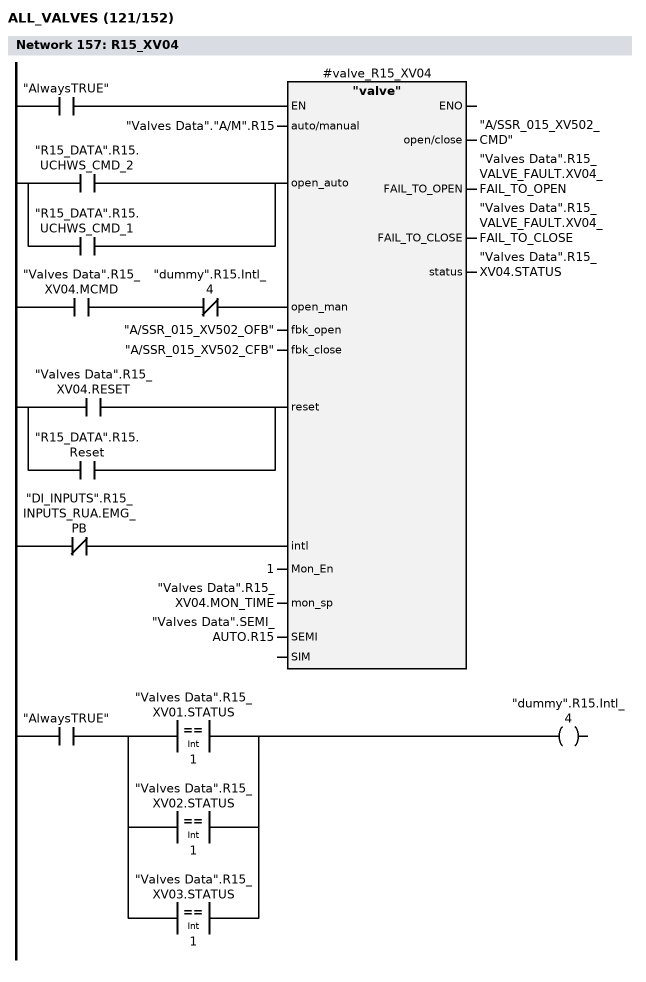
   RUNG wire#powerrail
      Contact( "AlwaysTRUE" )
      #valve_R15_XV04(open_auto := wire#w1, open_man := wire#w2, reset := wire#w3, intl := wire#w4, "auto/manual" := "Valves Data"."A/M".R15, fbk_open := "A/SSR_015_XV502_OFB", fbk_close := "A/SSR_015_XV502_CFB", Mon_En := 1, mon_sp := "Valves Data".R15_XV04.MON_TIME, SEMI := "Valves Data".SEMI_AUTO.R15, SIM :=, "open/close" => "A/SSR_015_XV502_CMD", FAIL_TO_OPEN => "Valves Data".R15_VALVE_FAULT.XV04_FAIL_TO_OPEN, FAIL_TO_CLOSE => "Valves Data".R15_VALVE_FAULT.XV04_FAIL_TO_CLOSE, status => "Valves Data".R15_XV04.STATUS)
   END_RUNG
   RUNG wire#powerrail
      Contact( "R15_DATA".R15.UCHWS_CMD_2 )
   END_RUNG wire#w1
   RUNG wire#powerrail
      Contact( "R15_DATA".R15.UCHWS_CMD_1 )
   END_RUNG wire#w1
   RUNG wire#powerrail
      Contact( "Valves Data".R15_XV04.MCMD )
      I_Contact( "dummy".R15.Intl_4 )
   END_RUNG wire#w2
   RUNG wire#powerrail
      Contact( "Valves Data".R15_XV04.RESET )
   END_RUNG wire#w3
   RUNG wire#powerrail
      Contact( "R15_DATA".R15.Reset )
   END_RUNG wire#w3
   RUNG wire#powerrail
      I_Contact( "DI_INPUTS".R15_INPUTS_RUA.EMG_PB )
   END_RUNG wire#w4
   RUNG wire#powerrail
      Contact( "AlwaysTRUE" )
      wire#w5
      { S7_Templates := "SrcType := Int" } EQ_Contact(in1 := "Valves Data".R15_XV01.STATUS, in2 := 1)
      wire#w6
      Coil( "dummy".R15.Intl_4 )
   END_RUNG
   RUNG wire#w5
      { S7_Templates := "SrcType := Int" } EQ_Contact(in1 := "Valves Data".R15_XV02.STATUS, in2 := 1)
   END_RUNG wire#w6
   RUNG wire#w5
      { S7_Templates := "SrcType := Int" } EQ_Contact(in1 := "Valves Data".R15_XV03.STATUS, in2 := 1)
   END_RUNG wire#w6
   // the same network as SCL:
   IF "AlwaysTRUE" THEN
       #valve_R15_XV04("auto/manual" := "Valves Data"."A/M".R15,   // "valve"
                       open_auto := "R15_DATA".R15.UCHWS_CMD_2 OR "R15_DATA".R15.UCHWS_CMD_1,
                       open_man := "Valves Data".R15_XV04.MCMD AND NOT "dummy".R15.Intl_4,
                       fbk_open := "A/SSR_015_XV502_OFB",
                       fbk_close := "A/SSR_015_XV502_CFB",
                       reset := "Valves Data".R15_XV04.RESET OR "R15_DATA".R15.Reset,
                       intl := NOT "DI_INPUTS".R15_INPUTS_RUA.EMG_PB,
                       Mon_En := 1,
                       mon_sp := "Valves Data".R15_XV04.MON_TIME,
                       SEMI := "Valves Data".SEMI_AUTO.R15,
                       "open/close" => "A/SSR_015_XV502_CMD",
                       FAIL_TO_OPEN => "Valves Data".R15_VALVE_FAULT.XV04_FAIL_TO_OPEN,
                       FAIL_TO_CLOSE => "Valves Data".R15_VALVE_FAULT.XV04_FAIL_TO_CLOSE,
                       status => "Valves Data".R15_XV04.STATUS);
   END_IF;
   "dummy".R15.Intl_4 := "AlwaysTRUE" AND (("Valves Data".R15_XV01.STATUS = 1) OR ("Valves Data".R15_XV02.STATUS = 1) OR ("Valves Data".R15_XV03.STATUS = 1));
END_REGION

REGION Network 158: R15_XV05
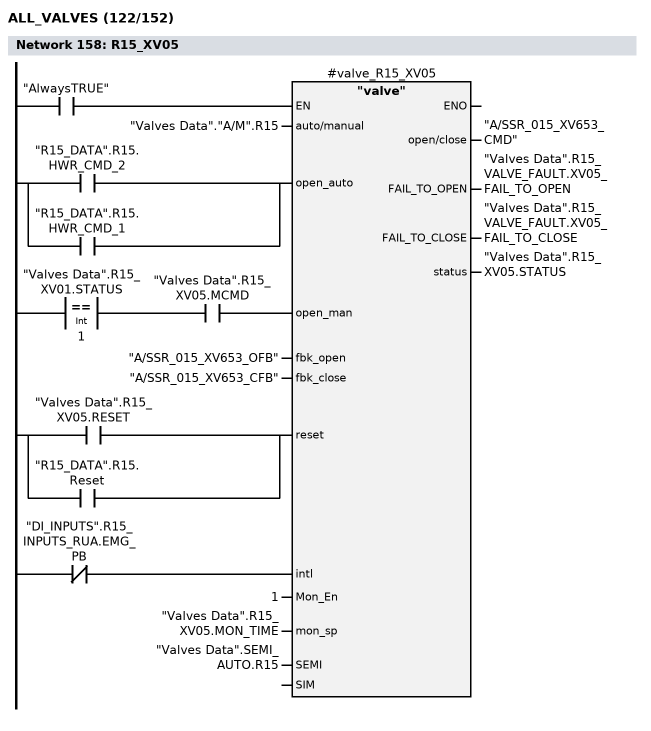
   RUNG wire#powerrail
      Contact( "AlwaysTRUE" )
      #valve_R15_XV05(open_auto := wire#w1, open_man := wire#w2, reset := wire#w3, intl := wire#w4, "auto/manual" := "Valves Data"."A/M".R15, fbk_open := "A/SSR_015_XV653_OFB", fbk_close := "A/SSR_015_XV653_CFB", Mon_En := 1, mon_sp := "Valves Data".R15_XV05.MON_TIME, SEMI := "Valves Data".SEMI_AUTO.R15, SIM :=, "open/close" => "A/SSR_015_XV653_CMD", FAIL_TO_OPEN => "Valves Data".R15_VALVE_FAULT.XV05_FAIL_TO_OPEN, FAIL_TO_CLOSE => "Valves Data".R15_VALVE_FAULT.XV05_FAIL_TO_CLOSE, status => "Valves Data".R15_XV05.STATUS)
   END_RUNG
   RUNG wire#powerrail
      Contact( "R15_DATA".R15.HWR_CMD_2 )
   END_RUNG wire#w1
   RUNG wire#powerrail
      Contact( "R15_DATA".R15.HWR_CMD_1 )
   END_RUNG wire#w1
   RUNG wire#powerrail
      { S7_Templates := "SrcType := Int" } EQ_Contact(in1 := "Valves Data".R15_XV01.STATUS, in2 := 1)
      Contact( "Valves Data".R15_XV05.MCMD )
   END_RUNG wire#w2
   RUNG wire#powerrail
      Contact( "Valves Data".R15_XV05.RESET )
   END_RUNG wire#w3
   RUNG wire#powerrail
      Contact( "R15_DATA".R15.Reset )
   END_RUNG wire#w3
   RUNG wire#powerrail
      I_Contact( "DI_INPUTS".R15_INPUTS_RUA.EMG_PB )
   END_RUNG wire#w4
   // the same network as SCL:
   IF "AlwaysTRUE" THEN
       #valve_R15_XV05("auto/manual" := "Valves Data"."A/M".R15,   // "valve"
                       open_auto := "R15_DATA".R15.HWR_CMD_2 OR "R15_DATA".R15.HWR_CMD_1,
                       open_man := ("Valves Data".R15_XV01.STATUS = 1) AND "Valves Data".R15_XV05.MCMD,
                       fbk_open := "A/SSR_015_XV653_OFB",
                       fbk_close := "A/SSR_015_XV653_CFB",
                       reset := "Valves Data".R15_XV05.RESET OR "R15_DATA".R15.Reset,
                       intl := NOT "DI_INPUTS".R15_INPUTS_RUA.EMG_PB,
                       Mon_En := 1,
                       mon_sp := "Valves Data".R15_XV05.MON_TIME,
                       SEMI := "Valves Data".SEMI_AUTO.R15,
                       "open/close" => "A/SSR_015_XV653_CMD",
                       FAIL_TO_OPEN => "Valves Data".R15_VALVE_FAULT.XV05_FAIL_TO_OPEN,
                       FAIL_TO_CLOSE => "Valves Data".R15_VALVE_FAULT.XV05_FAIL_TO_CLOSE,
                       status => "Valves Data".R15_XV05.STATUS);
   END_IF;
END_REGION

REGION Network 159: R15_XV06
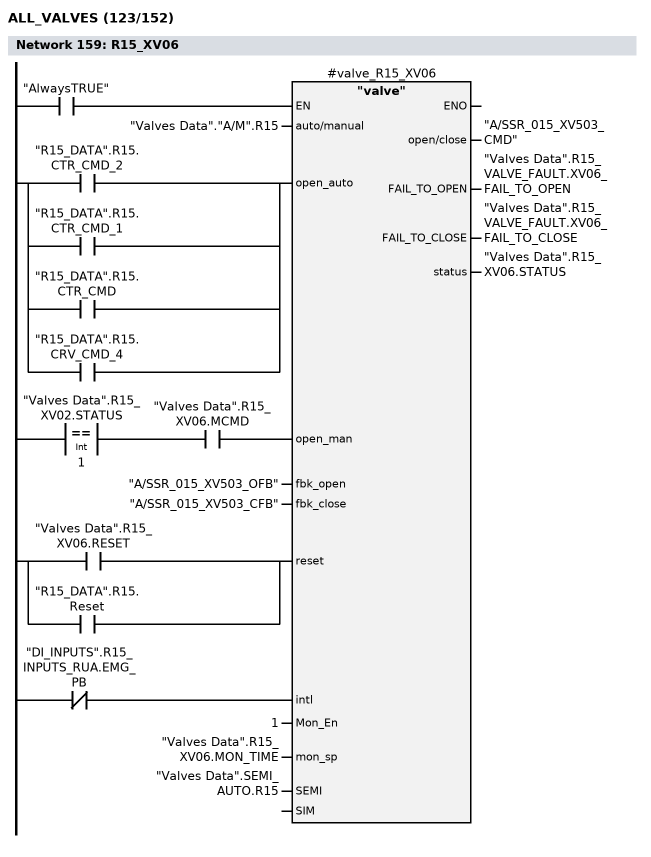
   RUNG wire#powerrail
      Contact( "AlwaysTRUE" )
      #valve_R15_XV06(open_auto := wire#w1, open_man := wire#w2, reset := wire#w3, intl := wire#w4, "auto/manual" := "Valves Data"."A/M".R15, fbk_open := "A/SSR_015_XV503_OFB", fbk_close := "A/SSR_015_XV503_CFB", Mon_En := 1, mon_sp := "Valves Data".R15_XV06.MON_TIME, SEMI := "Valves Data".SEMI_AUTO.R15, SIM :=, "open/close" => "A/SSR_015_XV503_CMD", FAIL_TO_OPEN => "Valves Data".R15_VALVE_FAULT.XV06_FAIL_TO_OPEN, FAIL_TO_CLOSE => "Valves Data".R15_VALVE_FAULT.XV06_FAIL_TO_CLOSE, status => "Valves Data".R15_XV06.STATUS)
   END_RUNG
   RUNG wire#powerrail
      Contact( "R15_DATA".R15.CTR_CMD_2 )
   END_RUNG wire#w1
   RUNG wire#powerrail
      Contact( "R15_DATA".R15.CTR_CMD_1 )
   END_RUNG wire#w1
   RUNG wire#powerrail
      Contact( "R15_DATA".R15.CTR_CMD )
   END_RUNG wire#w1
   RUNG wire#powerrail
      Contact( "R15_DATA".R15.CRV_CMD_4 )
   END_RUNG wire#w1
   RUNG wire#powerrail
      { S7_Templates := "SrcType := Int" } EQ_Contact(in1 := "Valves Data".R15_XV02.STATUS, in2 := 1)
      Contact( "Valves Data".R15_XV06.MCMD )
   END_RUNG wire#w2
   RUNG wire#powerrail
      Contact( "Valves Data".R15_XV06.RESET )
   END_RUNG wire#w3
   RUNG wire#powerrail
      Contact( "R15_DATA".R15.Reset )
   END_RUNG wire#w3
   RUNG wire#powerrail
      I_Contact( "DI_INPUTS".R15_INPUTS_RUA.EMG_PB )
   END_RUNG wire#w4
   // the same network as SCL:
   IF "AlwaysTRUE" THEN
       #valve_R15_XV06("auto/manual" := "Valves Data"."A/M".R15,   // "valve"
                       open_auto := "R15_DATA".R15.CTR_CMD_2 OR "R15_DATA".R15.CTR_CMD_1 OR "R15_DATA".R15.CTR_CMD OR "R15_DATA".R15.CRV_CMD_4,
                       open_man := ("Valves Data".R15_XV02.STATUS = 1) AND "Valves Data".R15_XV06.MCMD,
                       fbk_open := "A/SSR_015_XV503_OFB",
                       fbk_close := "A/SSR_015_XV503_CFB",
                       reset := "Valves Data".R15_XV06.RESET OR "R15_DATA".R15.Reset,
                       intl := NOT "DI_INPUTS".R15_INPUTS_RUA.EMG_PB,
                       Mon_En := 1,
                       mon_sp := "Valves Data".R15_XV06.MON_TIME,
                       SEMI := "Valves Data".SEMI_AUTO.R15,
                       "open/close" => "A/SSR_015_XV503_CMD",
                       FAIL_TO_OPEN => "Valves Data".R15_VALVE_FAULT.XV06_FAIL_TO_OPEN,
                       FAIL_TO_CLOSE => "Valves Data".R15_VALVE_FAULT.XV06_FAIL_TO_CLOSE,
                       status => "Valves Data".R15_XV06.STATUS);
   END_IF;
END_REGION

REGION Network 160: R15_XV07
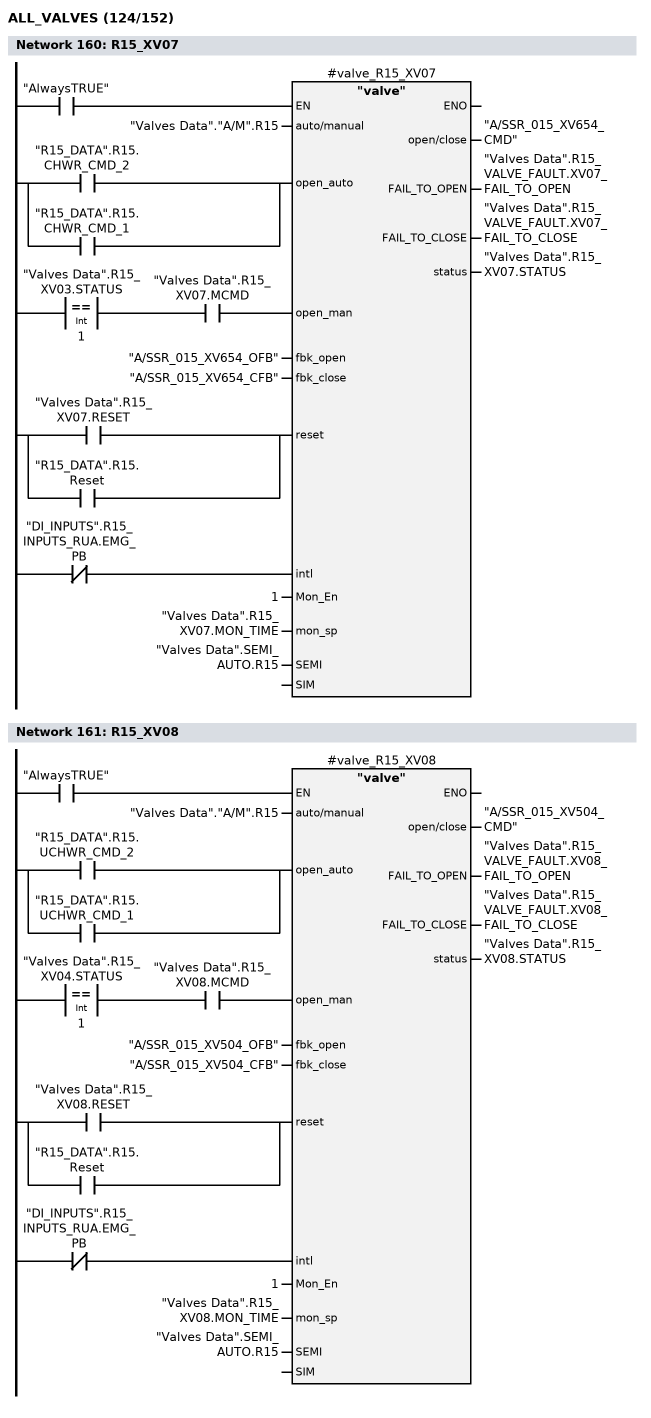
   RUNG wire#powerrail
      Contact( "AlwaysTRUE" )
      #valve_R15_XV07(open_auto := wire#w1, open_man := wire#w2, reset := wire#w3, intl := wire#w4, "auto/manual" := "Valves Data"."A/M".R15, fbk_open := "A/SSR_015_XV654_OFB", fbk_close := "A/SSR_015_XV654_CFB", Mon_En := 1, mon_sp := "Valves Data".R15_XV07.MON_TIME, SEMI := "Valves Data".SEMI_AUTO.R15, SIM :=, "open/close" => "A/SSR_015_XV654_CMD", FAIL_TO_OPEN => "Valves Data".R15_VALVE_FAULT.XV07_FAIL_TO_OPEN, FAIL_TO_CLOSE => "Valves Data".R15_VALVE_FAULT.XV07_FAIL_TO_CLOSE, status => "Valves Data".R15_XV07.STATUS)
   END_RUNG
   RUNG wire#powerrail
      Contact( "R15_DATA".R15.CHWR_CMD_2 )
   END_RUNG wire#w1
   RUNG wire#powerrail
      Contact( "R15_DATA".R15.CHWR_CMD_1 )
   END_RUNG wire#w1
   RUNG wire#powerrail
      { S7_Templates := "SrcType := Int" } EQ_Contact(in1 := "Valves Data".R15_XV03.STATUS, in2 := 1)
      Contact( "Valves Data".R15_XV07.MCMD )
   END_RUNG wire#w2
   RUNG wire#powerrail
      Contact( "Valves Data".R15_XV07.RESET )
   END_RUNG wire#w3
   RUNG wire#powerrail
      Contact( "R15_DATA".R15.Reset )
   END_RUNG wire#w3
   RUNG wire#powerrail
      I_Contact( "DI_INPUTS".R15_INPUTS_RUA.EMG_PB )
   END_RUNG wire#w4
   // the same network as SCL:
   IF "AlwaysTRUE" THEN
       #valve_R15_XV07("auto/manual" := "Valves Data"."A/M".R15,   // "valve"
                       open_auto := "R15_DATA".R15.CHWR_CMD_2 OR "R15_DATA".R15.CHWR_CMD_1,
                       open_man := ("Valves Data".R15_XV03.STATUS = 1) AND "Valves Data".R15_XV07.MCMD,
                       fbk_open := "A/SSR_015_XV654_OFB",
                       fbk_close := "A/SSR_015_XV654_CFB",
                       reset := "Valves Data".R15_XV07.RESET OR "R15_DATA".R15.Reset,
                       intl := NOT "DI_INPUTS".R15_INPUTS_RUA.EMG_PB,
                       Mon_En := 1,
                       mon_sp := "Valves Data".R15_XV07.MON_TIME,
                       SEMI := "Valves Data".SEMI_AUTO.R15,
                       "open/close" => "A/SSR_015_XV654_CMD",
                       FAIL_TO_OPEN => "Valves Data".R15_VALVE_FAULT.XV07_FAIL_TO_OPEN,
                       FAIL_TO_CLOSE => "Valves Data".R15_VALVE_FAULT.XV07_FAIL_TO_CLOSE,
                       status => "Valves Data".R15_XV07.STATUS);
   END_IF;
END_REGION

REGION Network 161: R15_XV08
   RUNG wire#powerrail
      Contact( "AlwaysTRUE" )
      #valve_R15_XV08(open_auto := wire#w1, open_man := wire#w2, reset := wire#w3, intl := wire#w4, "auto/manual" := "Valves Data"."A/M".R15, fbk_open := "A/SSR_015_XV504_OFB", fbk_close := "A/SSR_015_XV504_CFB", Mon_En := 1, mon_sp := "Valves Data".R15_XV08.MON_TIME, SEMI := "Valves Data".SEMI_AUTO.R15, SIM :=, "open/close" => "A/SSR_015_XV504_CMD", FAIL_TO_OPEN => "Valves Data".R15_VALVE_FAULT.XV08_FAIL_TO_OPEN, FAIL_TO_CLOSE => "Valves Data".R15_VALVE_FAULT.XV08_FAIL_TO_CLOSE, status => "Valves Data".R15_XV08.STATUS)
   END_RUNG
   RUNG wire#powerrail
      Contact( "R15_DATA".R15.UCHWR_CMD_2 )
   END_RUNG wire#w1
   RUNG wire#powerrail
      Contact( "R15_DATA".R15.UCHWR_CMD_1 )
   END_RUNG wire#w1
   RUNG wire#powerrail
      { S7_Templates := "SrcType := Int" } EQ_Contact(in1 := "Valves Data".R15_XV04.STATUS, in2 := 1)
      Contact( "Valves Data".R15_XV08.MCMD )
   END_RUNG wire#w2
   RUNG wire#powerrail
      Contact( "Valves Data".R15_XV08.RESET )
   END_RUNG wire#w3
   RUNG wire#powerrail
      Contact( "R15_DATA".R15.Reset )
   END_RUNG wire#w3
   RUNG wire#powerrail
      I_Contact( "DI_INPUTS".R15_INPUTS_RUA.EMG_PB )
   END_RUNG wire#w4
   // the same network as SCL:
   IF "AlwaysTRUE" THEN
       #valve_R15_XV08("auto/manual" := "Valves Data"."A/M".R15,   // "valve"
                       open_auto := "R15_DATA".R15.UCHWR_CMD_2 OR "R15_DATA".R15.UCHWR_CMD_1,
                       open_man := ("Valves Data".R15_XV04.STATUS = 1) AND "Valves Data".R15_XV08.MCMD,
                       fbk_open := "A/SSR_015_XV504_OFB",
                       fbk_close := "A/SSR_015_XV504_CFB",
                       reset := "Valves Data".R15_XV08.RESET OR "R15_DATA".R15.Reset,
                       intl := NOT "DI_INPUTS".R15_INPUTS_RUA.EMG_PB,
                       Mon_En := 1,
                       mon_sp := "Valves Data".R15_XV08.MON_TIME,
                       SEMI := "Valves Data".SEMI_AUTO.R15,
                       "open/close" => "A/SSR_015_XV504_CMD",
                       FAIL_TO_OPEN => "Valves Data".R15_VALVE_FAULT.XV08_FAIL_TO_OPEN,
                       FAIL_TO_CLOSE => "Valves Data".R15_VALVE_FAULT.XV08_FAIL_TO_CLOSE,
                       status => "Valves Data".R15_XV08.STATUS);
   END_IF;
END_REGION

REGION Network 162: R15_XV09
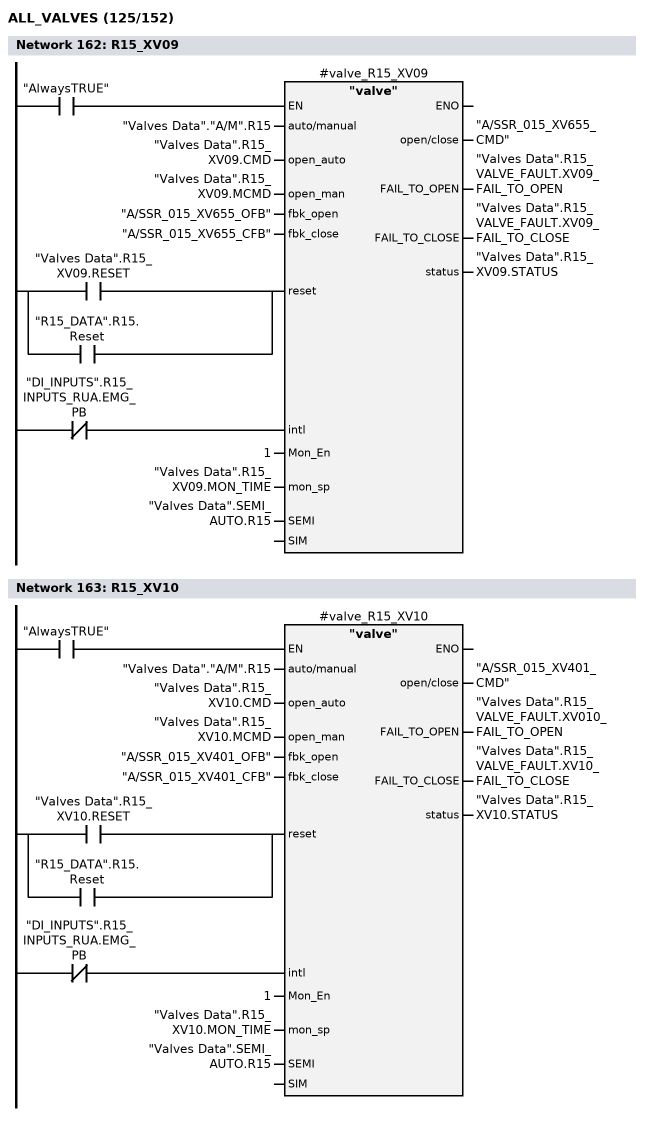
   RUNG wire#powerrail
      Contact( "AlwaysTRUE" )
      #valve_R15_XV09(reset := wire#w1, intl := wire#w2, "auto/manual" := "Valves Data"."A/M".R15, open_auto := "Valves Data".R15_XV09.CMD, open_man := "Valves Data".R15_XV09.MCMD, fbk_open := "A/SSR_015_XV655_OFB", fbk_close := "A/SSR_015_XV655_CFB", Mon_En := 1, mon_sp := "Valves Data".R15_XV09.MON_TIME, SEMI := "Valves Data".SEMI_AUTO.R15, SIM :=, "open/close" => "A/SSR_015_XV655_CMD", FAIL_TO_OPEN => "Valves Data".R15_VALVE_FAULT.XV09_FAIL_TO_OPEN, FAIL_TO_CLOSE => "Valves Data".R15_VALVE_FAULT.XV09_FAIL_TO_CLOSE, status => "Valves Data".R15_XV09.STATUS)
   END_RUNG
   RUNG wire#powerrail
      Contact( "Valves Data".R15_XV09.RESET )
   END_RUNG wire#w1
   RUNG wire#powerrail
      Contact( "R15_DATA".R15.Reset )
   END_RUNG wire#w1
   RUNG wire#powerrail
      I_Contact( "DI_INPUTS".R15_INPUTS_RUA.EMG_PB )
   END_RUNG wire#w2
   // the same network as SCL:
   IF "AlwaysTRUE" THEN
       #valve_R15_XV09("auto/manual" := "Valves Data"."A/M".R15,   // "valve"
                       open_auto := "Valves Data".R15_XV09.CMD,
                       open_man := "Valves Data".R15_XV09.MCMD,
                       fbk_open := "A/SSR_015_XV655_OFB",
                       fbk_close := "A/SSR_015_XV655_CFB",
                       reset := "Valves Data".R15_XV09.RESET OR "R15_DATA".R15.Reset,
                       intl := NOT "DI_INPUTS".R15_INPUTS_RUA.EMG_PB,
                       Mon_En := 1,
                       mon_sp := "Valves Data".R15_XV09.MON_TIME,
                       SEMI := "Valves Data".SEMI_AUTO.R15,
                       "open/close" => "A/SSR_015_XV655_CMD",
                       FAIL_TO_OPEN => "Valves Data".R15_VALVE_FAULT.XV09_FAIL_TO_OPEN,
                       FAIL_TO_CLOSE => "Valves Data".R15_VALVE_FAULT.XV09_FAIL_TO_CLOSE,
                       status => "Valves Data".R15_XV09.STATUS);
   END_IF;
END_REGION

REGION Network 163: R15_XV10
   RUNG wire#powerrail
      Contact( "AlwaysTRUE" )
      #valve_R15_XV10(reset := wire#w1, intl := wire#w2, "auto/manual" := "Valves Data"."A/M".R15, open_auto := "Valves Data".R15_XV10.CMD, open_man := "Valves Data".R15_XV10.MCMD, fbk_open := "A/SSR_015_XV401_OFB", fbk_close := "A/SSR_015_XV401_CFB", Mon_En := 1, mon_sp := "Valves Data".R15_XV10.MON_TIME, SEMI := "Valves Data".SEMI_AUTO.R15, SIM :=, "open/close" => "A/SSR_015_XV401_CMD", FAIL_TO_OPEN => "Valves Data".R15_VALVE_FAULT.XV010_FAIL_TO_OPEN, FAIL_TO_CLOSE => "Valves Data".R15_VALVE_FAULT.XV10_FAIL_TO_CLOSE, status => "Valves Data".R15_XV10.STATUS)
   END_RUNG
   RUNG wire#powerrail
      Contact( "Valves Data".R15_XV10.RESET )
   END_RUNG wire#w1
   RUNG wire#powerrail
      Contact( "R15_DATA".R15.Reset )
   END_RUNG wire#w1
   RUNG wire#powerrail
      I_Contact( "DI_INPUTS".R15_INPUTS_RUA.EMG_PB )
   END_RUNG wire#w2
   // the same network as SCL:
   IF "AlwaysTRUE" THEN
       #valve_R15_XV10("auto/manual" := "Valves Data"."A/M".R15,   // "valve"
                       open_auto := "Valves Data".R15_XV10.CMD,
                       open_man := "Valves Data".R15_XV10.MCMD,
                       fbk_open := "A/SSR_015_XV401_OFB",
                       fbk_close := "A/SSR_015_XV401_CFB",
                       reset := "Valves Data".R15_XV10.RESET OR "R15_DATA".R15.Reset,
                       intl := NOT "DI_INPUTS".R15_INPUTS_RUA.EMG_PB,
                       Mon_En := 1,
                       mon_sp := "Valves Data".R15_XV10.MON_TIME,
                       SEMI := "Valves Data".SEMI_AUTO.R15,
                       "open/close" => "A/SSR_015_XV401_CMD",
                       FAIL_TO_OPEN => "Valves Data".R15_VALVE_FAULT.XV010_FAIL_TO_OPEN,
                       FAIL_TO_CLOSE => "Valves Data".R15_VALVE_FAULT.XV10_FAIL_TO_CLOSE,
                       status => "Valves Data".R15_XV10.STATUS);
   END_IF;
END_REGION

REGION Network 164: ****REACTOR_16****
END_REGION

REGION Network 165: R16_XV01
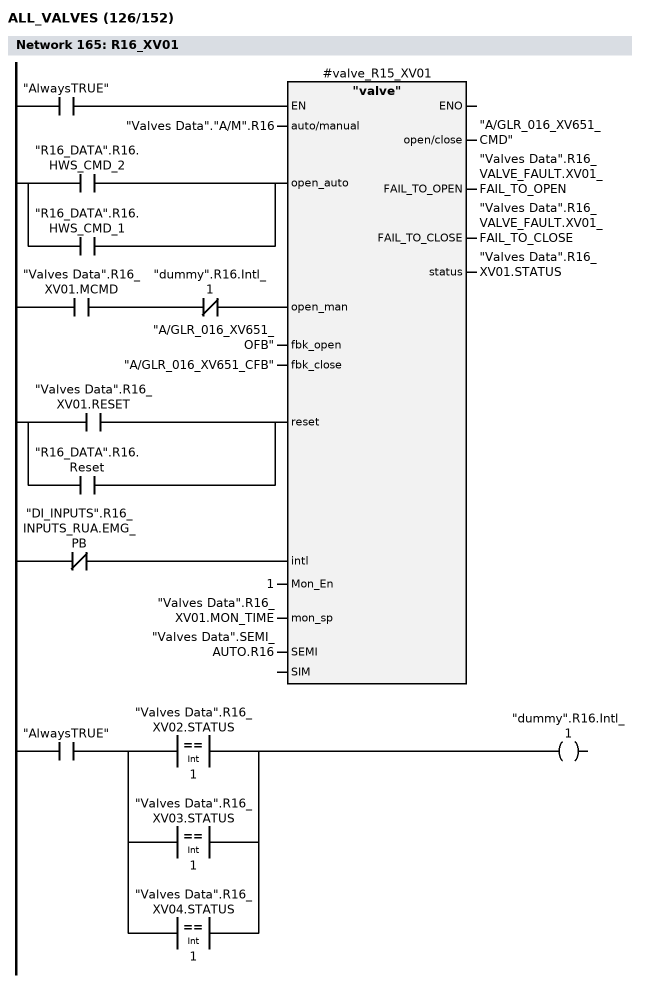
   RUNG wire#powerrail
      Contact( "AlwaysTRUE" )
      #valve_R15_XV01(open_auto := wire#w1, open_man := wire#w2, reset := wire#w3, intl := wire#w4, "auto/manual" := "Valves Data"."A/M".R16, fbk_open := "A/GLR_016_XV651_OFB", fbk_close := "A/GLR_016_XV651_CFB", Mon_En := 1, mon_sp := "Valves Data".R16_XV01.MON_TIME, SEMI := "Valves Data".SEMI_AUTO.R16, SIM :=, "open/close" => "A/GLR_016_XV651_CMD", FAIL_TO_OPEN => "Valves Data".R16_VALVE_FAULT.XV01_FAIL_TO_OPEN, FAIL_TO_CLOSE => "Valves Data".R16_VALVE_FAULT.XV01_FAIL_TO_CLOSE, status => "Valves Data".R16_XV01.STATUS)
   END_RUNG
   RUNG wire#powerrail
      Contact( "R16_DATA".R16.HWS_CMD_2 )
   END_RUNG wire#w1
   RUNG wire#powerrail
      Contact( "R16_DATA".R16.HWS_CMD_1 )
   END_RUNG wire#w1
   RUNG wire#powerrail
      Contact( "Valves Data".R16_XV01.MCMD )
      I_Contact( "dummy".R16.Intl_1 )
   END_RUNG wire#w2
   RUNG wire#powerrail
      Contact( "Valves Data".R16_XV01.RESET )
   END_RUNG wire#w3
   RUNG wire#powerrail
      Contact( "R16_DATA".R16.Reset )
   END_RUNG wire#w3
   RUNG wire#powerrail
      I_Contact( "DI_INPUTS".R16_INPUTS_RUA.EMG_PB )
   END_RUNG wire#w4
   RUNG wire#powerrail
      Contact( "AlwaysTRUE" )
      wire#w5
      { S7_Templates := "SrcType := Int" } EQ_Contact(in1 := "Valves Data".R16_XV02.STATUS, in2 := 1)
      wire#w6
      Coil( "dummy".R16.Intl_1 )
   END_RUNG
   RUNG wire#w5
      { S7_Templates := "SrcType := Int" } EQ_Contact(in1 := "Valves Data".R16_XV03.STATUS, in2 := 1)
   END_RUNG wire#w6
   RUNG wire#w5
      { S7_Templates := "SrcType := Int" } EQ_Contact(in1 := "Valves Data".R16_XV04.STATUS, in2 := 1)
   END_RUNG wire#w6
   // the same network as SCL:
   IF "AlwaysTRUE" THEN
       #valve_R15_XV01("auto/manual" := "Valves Data"."A/M".R16,   // "valve"
                       open_auto := "R16_DATA".R16.HWS_CMD_2 OR "R16_DATA".R16.HWS_CMD_1,
                       open_man := "Valves Data".R16_XV01.MCMD AND NOT "dummy".R16.Intl_1,
                       fbk_open := "A/GLR_016_XV651_OFB",
                       fbk_close := "A/GLR_016_XV651_CFB",
                       reset := "Valves Data".R16_XV01.RESET OR "R16_DATA".R16.Reset,
                       intl := NOT "DI_INPUTS".R16_INPUTS_RUA.EMG_PB,
                       Mon_En := 1,
                       mon_sp := "Valves Data".R16_XV01.MON_TIME,
                       SEMI := "Valves Data".SEMI_AUTO.R16,
                       "open/close" => "A/GLR_016_XV651_CMD",
                       FAIL_TO_OPEN => "Valves Data".R16_VALVE_FAULT.XV01_FAIL_TO_OPEN,
                       FAIL_TO_CLOSE => "Valves Data".R16_VALVE_FAULT.XV01_FAIL_TO_CLOSE,
                       status => "Valves Data".R16_XV01.STATUS);
   END_IF;
   "dummy".R16.Intl_1 := "AlwaysTRUE" AND (("Valves Data".R16_XV02.STATUS = 1) OR ("Valves Data".R16_XV03.STATUS = 1) OR ("Valves Data".R16_XV04.STATUS = 1));
END_REGION

REGION Network 166: R16_XV02
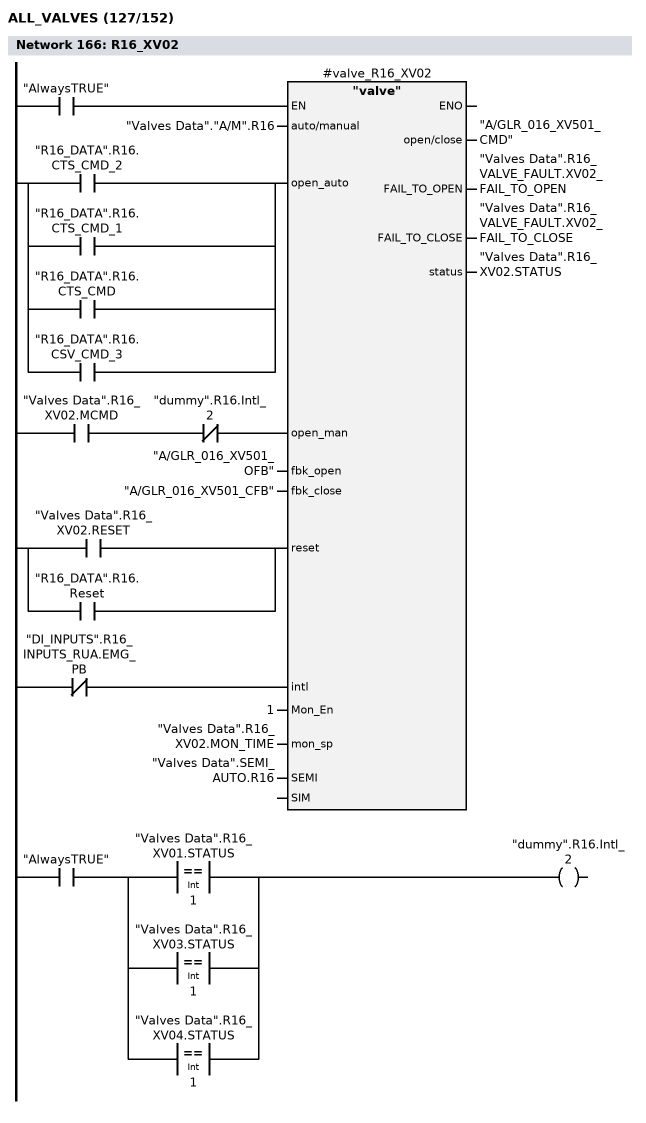
   RUNG wire#powerrail
      Contact( "AlwaysTRUE" )
      #valve_R16_XV02(open_auto := wire#w1, open_man := wire#w2, reset := wire#w3, intl := wire#w4, "auto/manual" := "Valves Data"."A/M".R16, fbk_open := "A/GLR_016_XV501_OFB", fbk_close := "A/GLR_016_XV501_CFB", Mon_En := 1, mon_sp := "Valves Data".R16_XV02.MON_TIME, SEMI := "Valves Data".SEMI_AUTO.R16, SIM :=, "open/close" => "A/GLR_016_XV501_CMD", FAIL_TO_OPEN => "Valves Data".R16_VALVE_FAULT.XV02_FAIL_TO_OPEN, FAIL_TO_CLOSE => "Valves Data".R16_VALVE_FAULT.XV02_FAIL_TO_CLOSE, status => "Valves Data".R16_XV02.STATUS)
   END_RUNG
   RUNG wire#powerrail
      Contact( "R16_DATA".R16.CTS_CMD_2 )
   END_RUNG wire#w1
   RUNG wire#powerrail
      Contact( "R16_DATA".R16.CTS_CMD_1 )
   END_RUNG wire#w1
   RUNG wire#powerrail
      Contact( "R16_DATA".R16.CTS_CMD )
   END_RUNG wire#w1
   RUNG wire#powerrail
      Contact( "R16_DATA".R16.CSV_CMD_3 )
   END_RUNG wire#w1
   RUNG wire#powerrail
      Contact( "Valves Data".R16_XV02.MCMD )
      I_Contact( "dummy".R16.Intl_2 )
   END_RUNG wire#w2
   RUNG wire#powerrail
      Contact( "Valves Data".R16_XV02.RESET )
   END_RUNG wire#w3
   RUNG wire#powerrail
      Contact( "R16_DATA".R16.Reset )
   END_RUNG wire#w3
   RUNG wire#powerrail
      I_Contact( "DI_INPUTS".R16_INPUTS_RUA.EMG_PB )
   END_RUNG wire#w4
   RUNG wire#powerrail
      Contact( "AlwaysTRUE" )
      wire#w5
      { S7_Templates := "SrcType := Int" } EQ_Contact(in1 := "Valves Data".R16_XV01.STATUS, in2 := 1)
      wire#w6
      Coil( "dummy".R16.Intl_2 )
   END_RUNG
   RUNG wire#w5
      { S7_Templates := "SrcType := Int" } EQ_Contact(in1 := "Valves Data".R16_XV03.STATUS, in2 := 1)
   END_RUNG wire#w6
   RUNG wire#w5
      { S7_Templates := "SrcType := Int" } EQ_Contact(in1 := "Valves Data".R16_XV04.STATUS, in2 := 1)
   END_RUNG wire#w6
   // the same network as SCL:
   IF "AlwaysTRUE" THEN
       #valve_R16_XV02("auto/manual" := "Valves Data"."A/M".R16,   // "valve"
                       open_auto := "R16_DATA".R16.CTS_CMD_2 OR "R16_DATA".R16.CTS_CMD_1 OR "R16_DATA".R16.CTS_CMD OR "R16_DATA".R16.CSV_CMD_3,
                       open_man := "Valves Data".R16_XV02.MCMD AND NOT "dummy".R16.Intl_2,
                       fbk_open := "A/GLR_016_XV501_OFB",
                       fbk_close := "A/GLR_016_XV501_CFB",
                       reset := "Valves Data".R16_XV02.RESET OR "R16_DATA".R16.Reset,
                       intl := NOT "DI_INPUTS".R16_INPUTS_RUA.EMG_PB,
                       Mon_En := 1,
                       mon_sp := "Valves Data".R16_XV02.MON_TIME,
                       SEMI := "Valves Data".SEMI_AUTO.R16,
                       "open/close" => "A/GLR_016_XV501_CMD",
                       FAIL_TO_OPEN => "Valves Data".R16_VALVE_FAULT.XV02_FAIL_TO_OPEN,
                       FAIL_TO_CLOSE => "Valves Data".R16_VALVE_FAULT.XV02_FAIL_TO_CLOSE,
                       status => "Valves Data".R16_XV02.STATUS);
   END_IF;
   "dummy".R16.Intl_2 := "AlwaysTRUE" AND (("Valves Data".R16_XV01.STATUS = 1) OR ("Valves Data".R16_XV03.STATUS = 1) OR ("Valves Data".R16_XV04.STATUS = 1));
END_REGION

REGION Network 167: R16_XV03
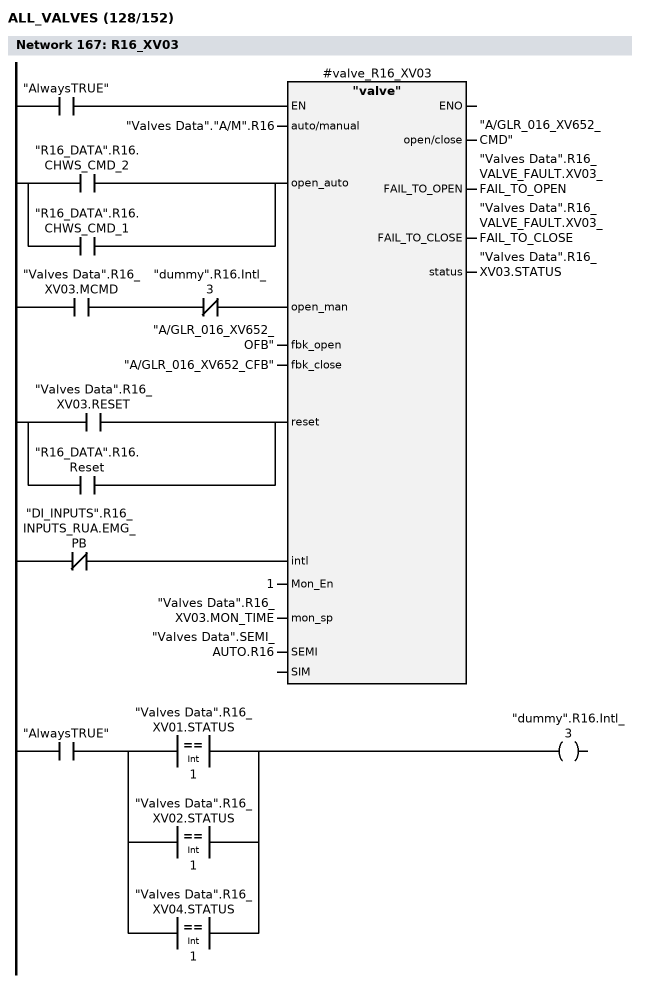
   RUNG wire#powerrail
      Contact( "AlwaysTRUE" )
      #valve_R16_XV03(open_auto := wire#w1, open_man := wire#w2, reset := wire#w3, intl := wire#w4, "auto/manual" := "Valves Data"."A/M".R16, fbk_open := "A/GLR_016_XV652_OFB", fbk_close := "A/GLR_016_XV652_CFB", Mon_En := 1, mon_sp := "Valves Data".R16_XV03.MON_TIME, SEMI := "Valves Data".SEMI_AUTO.R16, SIM :=, "open/close" => "A/GLR_016_XV652_CMD", FAIL_TO_OPEN => "Valves Data".R16_VALVE_FAULT.XV03_FAIL_TO_OPEN, FAIL_TO_CLOSE => "Valves Data".R16_VALVE_FAULT.XV03_FAIL_TO_CLOSE, status => "Valves Data".R16_XV03.STATUS)
   END_RUNG
   RUNG wire#powerrail
      Contact( "R16_DATA".R16.CHWS_CMD_2 )
   END_RUNG wire#w1
   RUNG wire#powerrail
      Contact( "R16_DATA".R16.CHWS_CMD_1 )
   END_RUNG wire#w1
   RUNG wire#powerrail
      Contact( "Valves Data".R16_XV03.MCMD )
      I_Contact( "dummy".R16.Intl_3 )
   END_RUNG wire#w2
   RUNG wire#powerrail
      Contact( "Valves Data".R16_XV03.RESET )
   END_RUNG wire#w3
   RUNG wire#powerrail
      Contact( "R16_DATA".R16.Reset )
   END_RUNG wire#w3
   RUNG wire#powerrail
      I_Contact( "DI_INPUTS".R16_INPUTS_RUA.EMG_PB )
   END_RUNG wire#w4
   RUNG wire#powerrail
      Contact( "AlwaysTRUE" )
      wire#w5
      { S7_Templates := "SrcType := Int" } EQ_Contact(in1 := "Valves Data".R16_XV01.STATUS, in2 := 1)
      wire#w6
      Coil( "dummy".R16.Intl_3 )
   END_RUNG
   RUNG wire#w5
      { S7_Templates := "SrcType := Int" } EQ_Contact(in1 := "Valves Data".R16_XV02.STATUS, in2 := 1)
   END_RUNG wire#w6
   RUNG wire#w5
      { S7_Templates := "SrcType := Int" } EQ_Contact(in1 := "Valves Data".R16_XV04.STATUS, in2 := 1)
   END_RUNG wire#w6
   // the same network as SCL:
   IF "AlwaysTRUE" THEN
       #valve_R16_XV03("auto/manual" := "Valves Data"."A/M".R16,   // "valve"
                       open_auto := "R16_DATA".R16.CHWS_CMD_2 OR "R16_DATA".R16.CHWS_CMD_1,
                       open_man := "Valves Data".R16_XV03.MCMD AND NOT "dummy".R16.Intl_3,
                       fbk_open := "A/GLR_016_XV652_OFB",
                       fbk_close := "A/GLR_016_XV652_CFB",
                       reset := "Valves Data".R16_XV03.RESET OR "R16_DATA".R16.Reset,
                       intl := NOT "DI_INPUTS".R16_INPUTS_RUA.EMG_PB,
                       Mon_En := 1,
                       mon_sp := "Valves Data".R16_XV03.MON_TIME,
                       SEMI := "Valves Data".SEMI_AUTO.R16,
                       "open/close" => "A/GLR_016_XV652_CMD",
                       FAIL_TO_OPEN => "Valves Data".R16_VALVE_FAULT.XV03_FAIL_TO_OPEN,
                       FAIL_TO_CLOSE => "Valves Data".R16_VALVE_FAULT.XV03_FAIL_TO_CLOSE,
                       status => "Valves Data".R16_XV03.STATUS);
   END_IF;
   "dummy".R16.Intl_3 := "AlwaysTRUE" AND (("Valves Data".R16_XV01.STATUS = 1) OR ("Valves Data".R16_XV02.STATUS = 1) OR ("Valves Data".R16_XV04.STATUS = 1));
END_REGION

REGION Network 168: R16_XV04
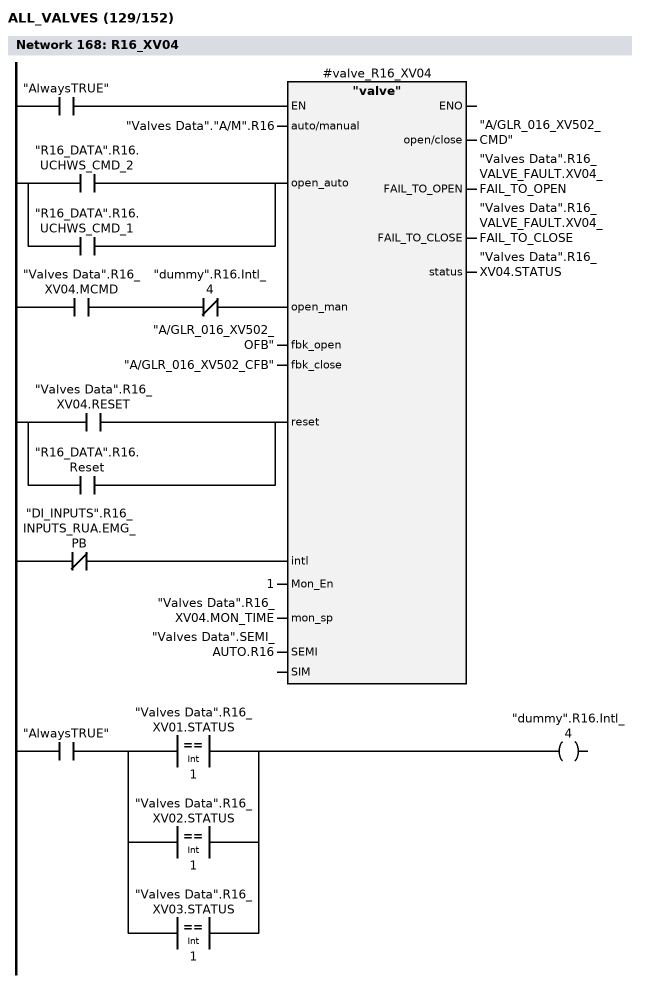
   RUNG wire#powerrail
      Contact( "AlwaysTRUE" )
      #valve_R16_XV04(open_auto := wire#w1, open_man := wire#w2, reset := wire#w3, intl := wire#w4, "auto/manual" := "Valves Data"."A/M".R16, fbk_open := "A/GLR_016_XV502_OFB", fbk_close := "A/GLR_016_XV502_CFB", Mon_En := 1, mon_sp := "Valves Data".R16_XV04.MON_TIME, SEMI := "Valves Data".SEMI_AUTO.R16, SIM :=, "open/close" => "A/GLR_016_XV502_CMD", FAIL_TO_OPEN => "Valves Data".R16_VALVE_FAULT.XV04_FAIL_TO_OPEN, FAIL_TO_CLOSE => "Valves Data".R16_VALVE_FAULT.XV04_FAIL_TO_CLOSE, status => "Valves Data".R16_XV04.STATUS)
   END_RUNG
   RUNG wire#powerrail
      Contact( "R16_DATA".R16.UCHWS_CMD_2 )
   END_RUNG wire#w1
   RUNG wire#powerrail
      Contact( "R16_DATA".R16.UCHWS_CMD_1 )
   END_RUNG wire#w1
   RUNG wire#powerrail
      Contact( "Valves Data".R16_XV04.MCMD )
      I_Contact( "dummy".R16.Intl_4 )
   END_RUNG wire#w2
   RUNG wire#powerrail
      Contact( "Valves Data".R16_XV04.RESET )
   END_RUNG wire#w3
   RUNG wire#powerrail
      Contact( "R16_DATA".R16.Reset )
   END_RUNG wire#w3
   RUNG wire#powerrail
      I_Contact( "DI_INPUTS".R16_INPUTS_RUA.EMG_PB )
   END_RUNG wire#w4
   RUNG wire#powerrail
      Contact( "AlwaysTRUE" )
      wire#w5
      { S7_Templates := "SrcType := Int" } EQ_Contact(in1 := "Valves Data".R16_XV01.STATUS, in2 := 1)
      wire#w6
      Coil( "dummy".R16.Intl_4 )
   END_RUNG
   RUNG wire#w5
      { S7_Templates := "SrcType := Int" } EQ_Contact(in1 := "Valves Data".R16_XV02.STATUS, in2 := 1)
   END_RUNG wire#w6
   RUNG wire#w5
      { S7_Templates := "SrcType := Int" } EQ_Contact(in1 := "Valves Data".R16_XV03.STATUS, in2 := 1)
   END_RUNG wire#w6
   // the same network as SCL:
   IF "AlwaysTRUE" THEN
       #valve_R16_XV04("auto/manual" := "Valves Data"."A/M".R16,   // "valve"
                       open_auto := "R16_DATA".R16.UCHWS_CMD_2 OR "R16_DATA".R16.UCHWS_CMD_1,
                       open_man := "Valves Data".R16_XV04.MCMD AND NOT "dummy".R16.Intl_4,
                       fbk_open := "A/GLR_016_XV502_OFB",
                       fbk_close := "A/GLR_016_XV502_CFB",
                       reset := "Valves Data".R16_XV04.RESET OR "R16_DATA".R16.Reset,
                       intl := NOT "DI_INPUTS".R16_INPUTS_RUA.EMG_PB,
                       Mon_En := 1,
                       mon_sp := "Valves Data".R16_XV04.MON_TIME,
                       SEMI := "Valves Data".SEMI_AUTO.R16,
                       "open/close" => "A/GLR_016_XV502_CMD",
                       FAIL_TO_OPEN => "Valves Data".R16_VALVE_FAULT.XV04_FAIL_TO_OPEN,
                       FAIL_TO_CLOSE => "Valves Data".R16_VALVE_FAULT.XV04_FAIL_TO_CLOSE,
                       status => "Valves Data".R16_XV04.STATUS);
   END_IF;
   "dummy".R16.Intl_4 := "AlwaysTRUE" AND (("Valves Data".R16_XV01.STATUS = 1) OR ("Valves Data".R16_XV02.STATUS = 1) OR ("Valves Data".R16_XV03.STATUS = 1));
END_REGION

REGION Network 169: R16_XV05
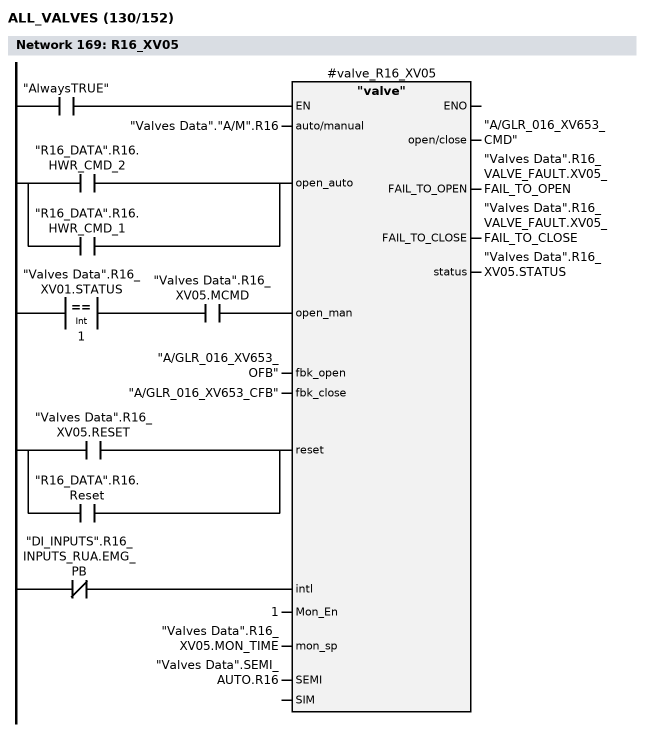
   RUNG wire#powerrail
      Contact( "AlwaysTRUE" )
      #valve_R16_XV05(open_auto := wire#w1, open_man := wire#w2, reset := wire#w3, intl := wire#w4, "auto/manual" := "Valves Data"."A/M".R16, fbk_open := "A/GLR_016_XV653_OFB", fbk_close := "A/GLR_016_XV653_CFB", Mon_En := 1, mon_sp := "Valves Data".R16_XV05.MON_TIME, SEMI := "Valves Data".SEMI_AUTO.R16, SIM :=, "open/close" => "A/GLR_016_XV653_CMD", FAIL_TO_OPEN => "Valves Data".R16_VALVE_FAULT.XV05_FAIL_TO_OPEN, FAIL_TO_CLOSE => "Valves Data".R16_VALVE_FAULT.XV05_FAIL_TO_CLOSE, status => "Valves Data".R16_XV05.STATUS)
   END_RUNG
   RUNG wire#powerrail
      Contact( "R16_DATA".R16.HWR_CMD_2 )
   END_RUNG wire#w1
   RUNG wire#powerrail
      Contact( "R16_DATA".R16.HWR_CMD_1 )
   END_RUNG wire#w1
   RUNG wire#powerrail
      { S7_Templates := "SrcType := Int" } EQ_Contact(in1 := "Valves Data".R16_XV01.STATUS, in2 := 1)
      Contact( "Valves Data".R16_XV05.MCMD )
   END_RUNG wire#w2
   RUNG wire#powerrail
      Contact( "Valves Data".R16_XV05.RESET )
   END_RUNG wire#w3
   RUNG wire#powerrail
      Contact( "R16_DATA".R16.Reset )
   END_RUNG wire#w3
   RUNG wire#powerrail
      I_Contact( "DI_INPUTS".R16_INPUTS_RUA.EMG_PB )
   END_RUNG wire#w4
   // the same network as SCL:
   IF "AlwaysTRUE" THEN
       #valve_R16_XV05("auto/manual" := "Valves Data"."A/M".R16,   // "valve"
                       open_auto := "R16_DATA".R16.HWR_CMD_2 OR "R16_DATA".R16.HWR_CMD_1,
                       open_man := ("Valves Data".R16_XV01.STATUS = 1) AND "Valves Data".R16_XV05.MCMD,
                       fbk_open := "A/GLR_016_XV653_OFB",
                       fbk_close := "A/GLR_016_XV653_CFB",
                       reset := "Valves Data".R16_XV05.RESET OR "R16_DATA".R16.Reset,
                       intl := NOT "DI_INPUTS".R16_INPUTS_RUA.EMG_PB,
                       Mon_En := 1,
                       mon_sp := "Valves Data".R16_XV05.MON_TIME,
                       SEMI := "Valves Data".SEMI_AUTO.R16,
                       "open/close" => "A/GLR_016_XV653_CMD",
                       FAIL_TO_OPEN => "Valves Data".R16_VALVE_FAULT.XV05_FAIL_TO_OPEN,
                       FAIL_TO_CLOSE => "Valves Data".R16_VALVE_FAULT.XV05_FAIL_TO_CLOSE,
                       status => "Valves Data".R16_XV05.STATUS);
   END_IF;
END_REGION

REGION Network 170: R16_XV06
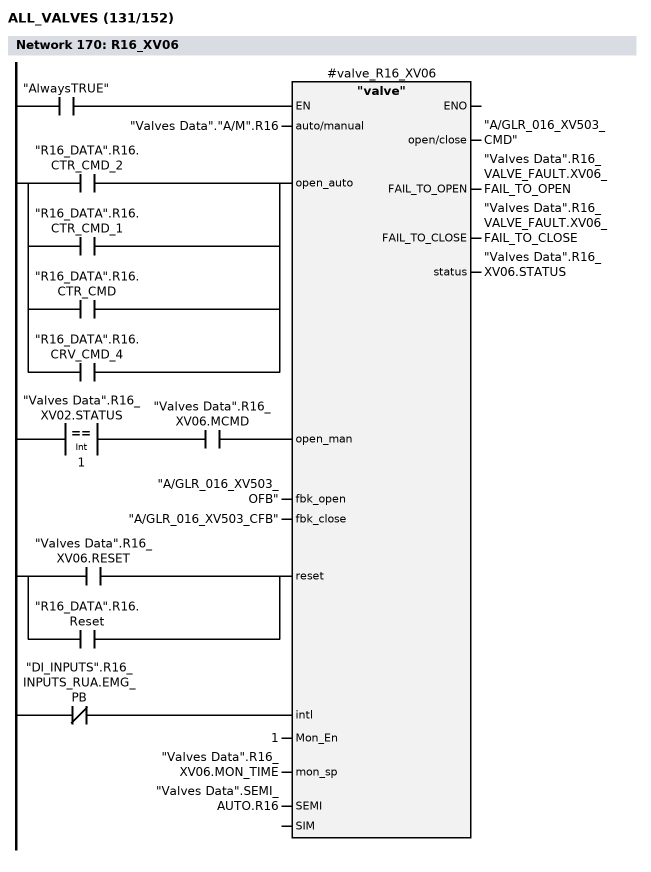
   RUNG wire#powerrail
      Contact( "AlwaysTRUE" )
      #valve_R16_XV06(open_auto := wire#w1, open_man := wire#w2, reset := wire#w3, intl := wire#w4, "auto/manual" := "Valves Data"."A/M".R16, fbk_open := "A/GLR_016_XV503_OFB", fbk_close := "A/GLR_016_XV503_CFB", Mon_En := 1, mon_sp := "Valves Data".R16_XV06.MON_TIME, SEMI := "Valves Data".SEMI_AUTO.R16, SIM :=, "open/close" => "A/GLR_016_XV503_CMD", FAIL_TO_OPEN => "Valves Data".R16_VALVE_FAULT.XV06_FAIL_TO_OPEN, FAIL_TO_CLOSE => "Valves Data".R16_VALVE_FAULT.XV06_FAIL_TO_CLOSE, status => "Valves Data".R16_XV06.STATUS)
   END_RUNG
   RUNG wire#powerrail
      Contact( "R16_DATA".R16.CTR_CMD_2 )
   END_RUNG wire#w1
   RUNG wire#powerrail
      Contact( "R16_DATA".R16.CTR_CMD_1 )
   END_RUNG wire#w1
   RUNG wire#powerrail
      Contact( "R16_DATA".R16.CTR_CMD )
   END_RUNG wire#w1
   RUNG wire#powerrail
      Contact( "R16_DATA".R16.CRV_CMD_4 )
   END_RUNG wire#w1
   RUNG wire#powerrail
      { S7_Templates := "SrcType := Int" } EQ_Contact(in1 := "Valves Data".R16_XV02.STATUS, in2 := 1)
      Contact( "Valves Data".R16_XV06.MCMD )
   END_RUNG wire#w2
   RUNG wire#powerrail
      Contact( "Valves Data".R16_XV06.RESET )
   END_RUNG wire#w3
   RUNG wire#powerrail
      Contact( "R16_DATA".R16.Reset )
   END_RUNG wire#w3
   RUNG wire#powerrail
      I_Contact( "DI_INPUTS".R16_INPUTS_RUA.EMG_PB )
   END_RUNG wire#w4
   // the same network as SCL:
   IF "AlwaysTRUE" THEN
       #valve_R16_XV06("auto/manual" := "Valves Data"."A/M".R16,   // "valve"
                       open_auto := "R16_DATA".R16.CTR_CMD_2 OR "R16_DATA".R16.CTR_CMD_1 OR "R16_DATA".R16.CTR_CMD OR "R16_DATA".R16.CRV_CMD_4,
                       open_man := ("Valves Data".R16_XV02.STATUS = 1) AND "Valves Data".R16_XV06.MCMD,
                       fbk_open := "A/GLR_016_XV503_OFB",
                       fbk_close := "A/GLR_016_XV503_CFB",
                       reset := "Valves Data".R16_XV06.RESET OR "R16_DATA".R16.Reset,
                       intl := NOT "DI_INPUTS".R16_INPUTS_RUA.EMG_PB,
                       Mon_En := 1,
                       mon_sp := "Valves Data".R16_XV06.MON_TIME,
                       SEMI := "Valves Data".SEMI_AUTO.R16,
                       "open/close" => "A/GLR_016_XV503_CMD",
                       FAIL_TO_OPEN => "Valves Data".R16_VALVE_FAULT.XV06_FAIL_TO_OPEN,
                       FAIL_TO_CLOSE => "Valves Data".R16_VALVE_FAULT.XV06_FAIL_TO_CLOSE,
                       status => "Valves Data".R16_XV06.STATUS);
   END_IF;
END_REGION

REGION Network 171: R16_XV07
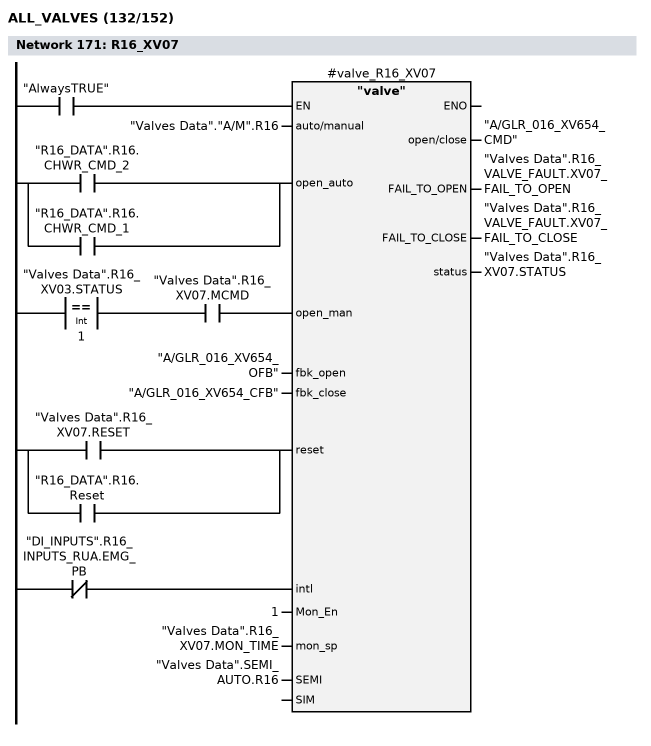
   RUNG wire#powerrail
      Contact( "AlwaysTRUE" )
      #valve_R16_XV07(open_auto := wire#w1, open_man := wire#w2, reset := wire#w3, intl := wire#w4, "auto/manual" := "Valves Data"."A/M".R16, fbk_open := "A/GLR_016_XV654_OFB", fbk_close := "A/GLR_016_XV654_CFB", Mon_En := 1, mon_sp := "Valves Data".R16_XV07.MON_TIME, SEMI := "Valves Data".SEMI_AUTO.R16, SIM :=, "open/close" => "A/GLR_016_XV654_CMD", FAIL_TO_OPEN => "Valves Data".R16_VALVE_FAULT.XV07_FAIL_TO_OPEN, FAIL_TO_CLOSE => "Valves Data".R16_VALVE_FAULT.XV07_FAIL_TO_CLOSE, status => "Valves Data".R16_XV07.STATUS)
   END_RUNG
   RUNG wire#powerrail
      Contact( "R16_DATA".R16.CHWR_CMD_2 )
   END_RUNG wire#w1
   RUNG wire#powerrail
      Contact( "R16_DATA".R16.CHWR_CMD_1 )
   END_RUNG wire#w1
   RUNG wire#powerrail
      { S7_Templates := "SrcType := Int" } EQ_Contact(in1 := "Valves Data".R16_XV03.STATUS, in2 := 1)
      Contact( "Valves Data".R16_XV07.MCMD )
   END_RUNG wire#w2
   RUNG wire#powerrail
      Contact( "Valves Data".R16_XV07.RESET )
   END_RUNG wire#w3
   RUNG wire#powerrail
      Contact( "R16_DATA".R16.Reset )
   END_RUNG wire#w3
   RUNG wire#powerrail
      I_Contact( "DI_INPUTS".R16_INPUTS_RUA.EMG_PB )
   END_RUNG wire#w4
   // the same network as SCL:
   IF "AlwaysTRUE" THEN
       #valve_R16_XV07("auto/manual" := "Valves Data"."A/M".R16,   // "valve"
                       open_auto := "R16_DATA".R16.CHWR_CMD_2 OR "R16_DATA".R16.CHWR_CMD_1,
                       open_man := ("Valves Data".R16_XV03.STATUS = 1) AND "Valves Data".R16_XV07.MCMD,
                       fbk_open := "A/GLR_016_XV654_OFB",
                       fbk_close := "A/GLR_016_XV654_CFB",
                       reset := "Valves Data".R16_XV07.RESET OR "R16_DATA".R16.Reset,
                       intl := NOT "DI_INPUTS".R16_INPUTS_RUA.EMG_PB,
                       Mon_En := 1,
                       mon_sp := "Valves Data".R16_XV07.MON_TIME,
                       SEMI := "Valves Data".SEMI_AUTO.R16,
                       "open/close" => "A/GLR_016_XV654_CMD",
                       FAIL_TO_OPEN => "Valves Data".R16_VALVE_FAULT.XV07_FAIL_TO_OPEN,
                       FAIL_TO_CLOSE => "Valves Data".R16_VALVE_FAULT.XV07_FAIL_TO_CLOSE,
                       status => "Valves Data".R16_XV07.STATUS);
   END_IF;
END_REGION

REGION Network 172: R16_XV08
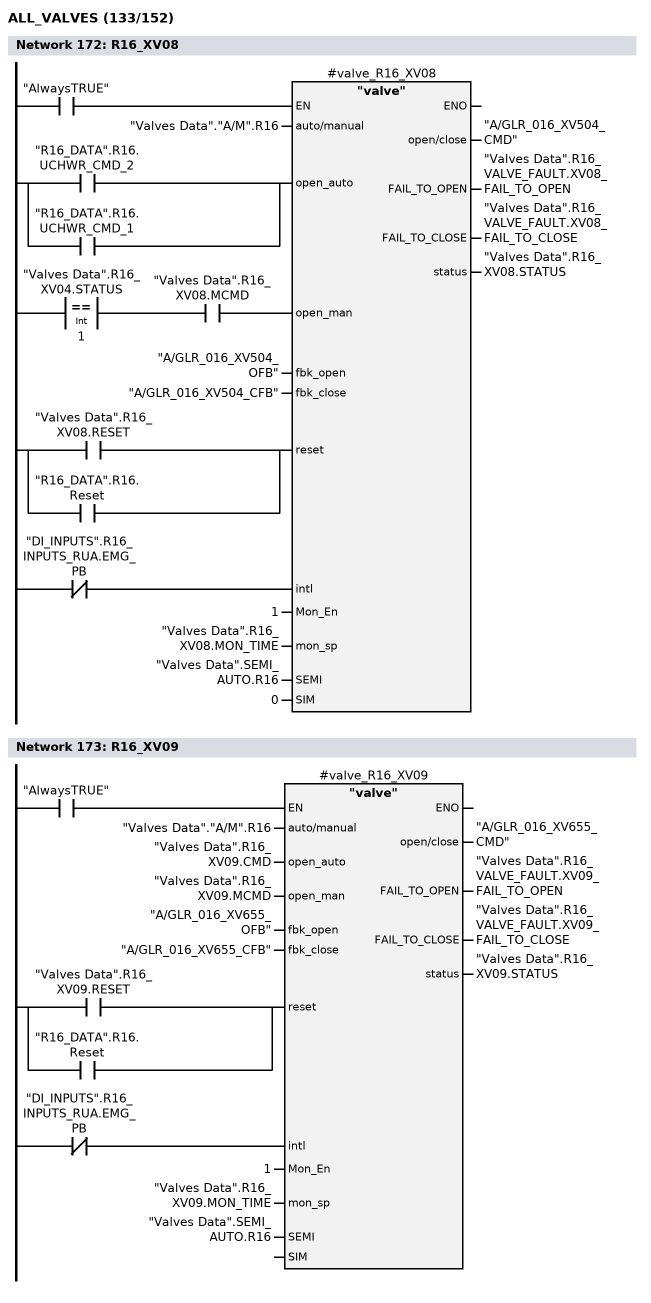
   RUNG wire#powerrail
      Contact( "AlwaysTRUE" )
      #valve_R16_XV08(open_auto := wire#w1, open_man := wire#w2, reset := wire#w3, intl := wire#w4, "auto/manual" := "Valves Data"."A/M".R16, fbk_open := "A/GLR_016_XV504_OFB", fbk_close := "A/GLR_016_XV504_CFB", Mon_En := 1, mon_sp := "Valves Data".R16_XV08.MON_TIME, SEMI := "Valves Data".SEMI_AUTO.R16, SIM := 0, "open/close" => "A/GLR_016_XV504_CMD", FAIL_TO_OPEN => "Valves Data".R16_VALVE_FAULT.XV08_FAIL_TO_OPEN, FAIL_TO_CLOSE => "Valves Data".R16_VALVE_FAULT.XV08_FAIL_TO_CLOSE, status => "Valves Data".R16_XV08.STATUS)
   END_RUNG
   RUNG wire#powerrail
      Contact( "R16_DATA".R16.UCHWR_CMD_2 )
   END_RUNG wire#w1
   RUNG wire#powerrail
      Contact( "R16_DATA".R16.UCHWR_CMD_1 )
   END_RUNG wire#w1
   RUNG wire#powerrail
      { S7_Templates := "SrcType := Int" } EQ_Contact(in1 := "Valves Data".R16_XV04.STATUS, in2 := 1)
      Contact( "Valves Data".R16_XV08.MCMD )
   END_RUNG wire#w2
   RUNG wire#powerrail
      Contact( "Valves Data".R16_XV08.RESET )
   END_RUNG wire#w3
   RUNG wire#powerrail
      Contact( "R16_DATA".R16.Reset )
   END_RUNG wire#w3
   RUNG wire#powerrail
      I_Contact( "DI_INPUTS".R16_INPUTS_RUA.EMG_PB )
   END_RUNG wire#w4
   // the same network as SCL:
   IF "AlwaysTRUE" THEN
       #valve_R16_XV08("auto/manual" := "Valves Data"."A/M".R16,   // "valve"
                       open_auto := "R16_DATA".R16.UCHWR_CMD_2 OR "R16_DATA".R16.UCHWR_CMD_1,
                       open_man := ("Valves Data".R16_XV04.STATUS = 1) AND "Valves Data".R16_XV08.MCMD,
                       fbk_open := "A/GLR_016_XV504_OFB",
                       fbk_close := "A/GLR_016_XV504_CFB",
                       reset := "Valves Data".R16_XV08.RESET OR "R16_DATA".R16.Reset,
                       intl := NOT "DI_INPUTS".R16_INPUTS_RUA.EMG_PB,
                       Mon_En := 1,
                       mon_sp := "Valves Data".R16_XV08.MON_TIME,
                       SEMI := "Valves Data".SEMI_AUTO.R16,
                       SIM := 0,
                       "open/close" => "A/GLR_016_XV504_CMD",
                       FAIL_TO_OPEN => "Valves Data".R16_VALVE_FAULT.XV08_FAIL_TO_OPEN,
                       FAIL_TO_CLOSE => "Valves Data".R16_VALVE_FAULT.XV08_FAIL_TO_CLOSE,
                       status => "Valves Data".R16_XV08.STATUS);
   END_IF;
END_REGION

REGION Network 173: R16_XV09
   RUNG wire#powerrail
      Contact( "AlwaysTRUE" )
      #valve_R16_XV09(reset := wire#w1, intl := wire#w2, "auto/manual" := "Valves Data"."A/M".R16, open_auto := "Valves Data".R16_XV09.CMD, open_man := "Valves Data".R16_XV09.MCMD, fbk_open := "A/GLR_016_XV655_OFB", fbk_close := "A/GLR_016_XV655_CFB", Mon_En := 1, mon_sp := "Valves Data".R16_XV09.MON_TIME, SEMI := "Valves Data".SEMI_AUTO.R16, SIM :=, "open/close" => "A/GLR_016_XV655_CMD", FAIL_TO_OPEN => "Valves Data".R16_VALVE_FAULT.XV09_FAIL_TO_OPEN, FAIL_TO_CLOSE => "Valves Data".R16_VALVE_FAULT.XV09_FAIL_TO_CLOSE, status => "Valves Data".R16_XV09.STATUS)
   END_RUNG
   RUNG wire#powerrail
      Contact( "Valves Data".R16_XV09.RESET )
   END_RUNG wire#w1
   RUNG wire#powerrail
      Contact( "R16_DATA".R16.Reset )
   END_RUNG wire#w1
   RUNG wire#powerrail
      I_Contact( "DI_INPUTS".R16_INPUTS_RUA.EMG_PB )
   END_RUNG wire#w2
   // the same network as SCL:
   IF "AlwaysTRUE" THEN
       #valve_R16_XV09("auto/manual" := "Valves Data"."A/M".R16,   // "valve"
                       open_auto := "Valves Data".R16_XV09.CMD,
                       open_man := "Valves Data".R16_XV09.MCMD,
                       fbk_open := "A/GLR_016_XV655_OFB",
                       fbk_close := "A/GLR_016_XV655_CFB",
                       reset := "Valves Data".R16_XV09.RESET OR "R16_DATA".R16.Reset,
                       intl := NOT "DI_INPUTS".R16_INPUTS_RUA.EMG_PB,
                       Mon_En := 1,
                       mon_sp := "Valves Data".R16_XV09.MON_TIME,
                       SEMI := "Valves Data".SEMI_AUTO.R16,
                       "open/close" => "A/GLR_016_XV655_CMD",
                       FAIL_TO_OPEN => "Valves Data".R16_VALVE_FAULT.XV09_FAIL_TO_OPEN,
                       FAIL_TO_CLOSE => "Valves Data".R16_VALVE_FAULT.XV09_FAIL_TO_CLOSE,
                       status => "Valves Data".R16_XV09.STATUS);
   END_IF;
END_REGION

REGION Network 174: R16_XV10
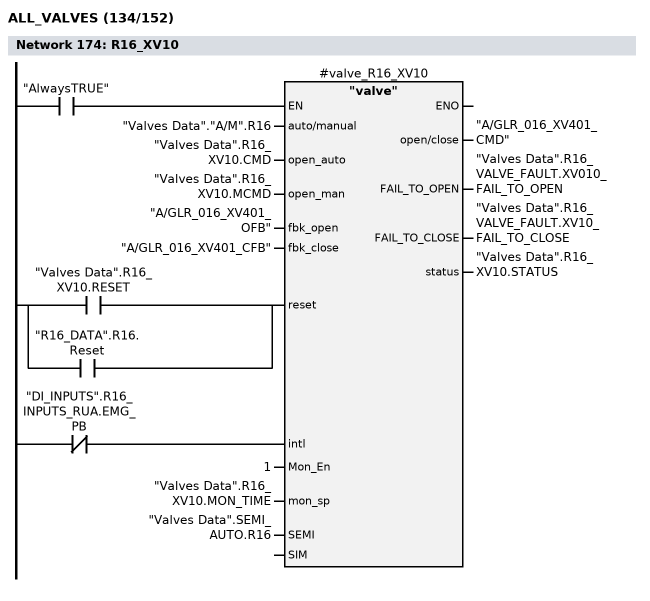
   RUNG wire#powerrail
      Contact( "AlwaysTRUE" )
      #valve_R16_XV10(reset := wire#w1, intl := wire#w2, "auto/manual" := "Valves Data"."A/M".R16, open_auto := "Valves Data".R16_XV10.CMD, open_man := "Valves Data".R16_XV10.MCMD, fbk_open := "A/GLR_016_XV401_OFB", fbk_close := "A/GLR_016_XV401_CFB", Mon_En := 1, mon_sp := "Valves Data".R16_XV10.MON_TIME, SEMI := "Valves Data".SEMI_AUTO.R16, SIM :=, "open/close" => "A/GLR_016_XV401_CMD", FAIL_TO_OPEN => "Valves Data".R16_VALVE_FAULT.XV010_FAIL_TO_OPEN, FAIL_TO_CLOSE => "Valves Data".R16_VALVE_FAULT.XV10_FAIL_TO_CLOSE, status => "Valves Data".R16_XV10.STATUS)
   END_RUNG
   RUNG wire#powerrail
      Contact( "Valves Data".R16_XV10.RESET )
   END_RUNG wire#w1
   RUNG wire#powerrail
      Contact( "R16_DATA".R16.Reset )
   END_RUNG wire#w1
   RUNG wire#powerrail
      I_Contact( "DI_INPUTS".R16_INPUTS_RUA.EMG_PB )
   END_RUNG wire#w2
   // the same network as SCL:
   IF "AlwaysTRUE" THEN
       #valve_R16_XV10("auto/manual" := "Valves Data"."A/M".R16,   // "valve"
                       open_auto := "Valves Data".R16_XV10.CMD,
                       open_man := "Valves Data".R16_XV10.MCMD,
                       fbk_open := "A/GLR_016_XV401_OFB",
                       fbk_close := "A/GLR_016_XV401_CFB",
                       reset := "Valves Data".R16_XV10.RESET OR "R16_DATA".R16.Reset,
                       intl := NOT "DI_INPUTS".R16_INPUTS_RUA.EMG_PB,
                       Mon_En := 1,
                       mon_sp := "Valves Data".R16_XV10.MON_TIME,
                       SEMI := "Valves Data".SEMI_AUTO.R16,
                       "open/close" => "A/GLR_016_XV401_CMD",
                       FAIL_TO_OPEN => "Valves Data".R16_VALVE_FAULT.XV010_FAIL_TO_OPEN,
                       FAIL_TO_CLOSE => "Valves Data".R16_VALVE_FAULT.XV10_FAIL_TO_CLOSE,
                       status => "Valves Data".R16_XV10.STATUS);
   END_IF;
END_REGION

REGION Network 175: ****REACTOR_17****
END_REGION

REGION Network 176: R17_XV01
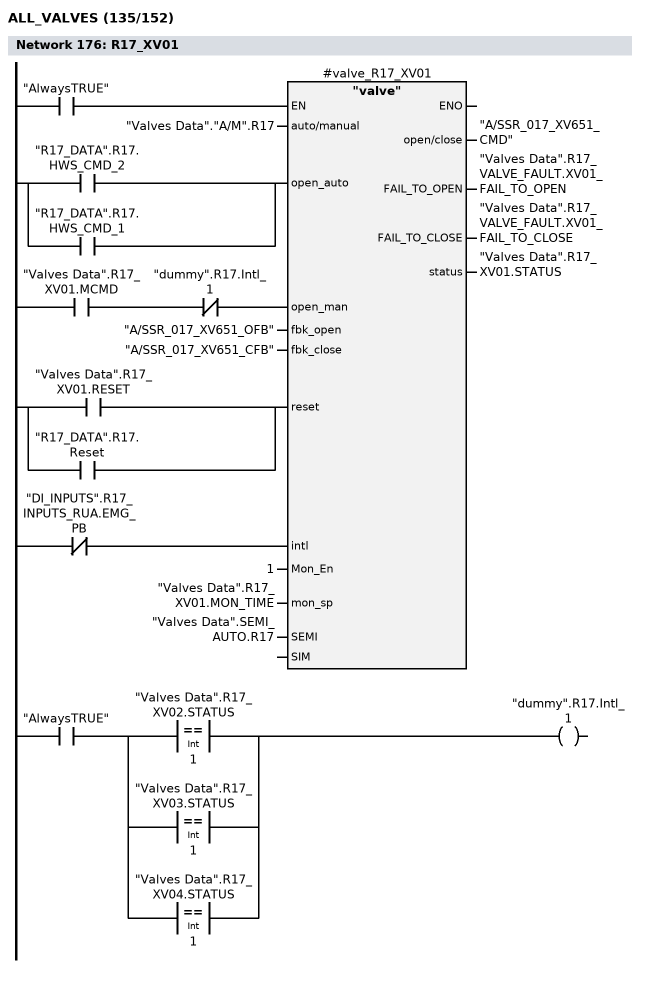
   RUNG wire#powerrail
      Contact( "AlwaysTRUE" )
      #valve_R17_XV01(open_auto := wire#w1, open_man := wire#w2, reset := wire#w3, intl := wire#w4, "auto/manual" := "Valves Data"."A/M".R17, fbk_open := "A/SSR_017_XV651_OFB", fbk_close := "A/SSR_017_XV651_CFB", Mon_En := 1, mon_sp := "Valves Data".R17_XV01.MON_TIME, SEMI := "Valves Data".SEMI_AUTO.R17, SIM :=, "open/close" => "A/SSR_017_XV651_CMD", FAIL_TO_OPEN => "Valves Data".R17_VALVE_FAULT.XV01_FAIL_TO_OPEN, FAIL_TO_CLOSE => "Valves Data".R17_VALVE_FAULT.XV01_FAIL_TO_CLOSE, status => "Valves Data".R17_XV01.STATUS)
   END_RUNG
   RUNG wire#powerrail
      Contact( "R17_DATA".R17.HWS_CMD_2 )
   END_RUNG wire#w1
   RUNG wire#powerrail
      Contact( "R17_DATA".R17.HWS_CMD_1 )
   END_RUNG wire#w1
   RUNG wire#powerrail
      Contact( "Valves Data".R17_XV01.MCMD )
      I_Contact( "dummy".R17.Intl_1 )
   END_RUNG wire#w2
   RUNG wire#powerrail
      Contact( "Valves Data".R17_XV01.RESET )
   END_RUNG wire#w3
   RUNG wire#powerrail
      Contact( "R17_DATA".R17.Reset )
   END_RUNG wire#w3
   RUNG wire#powerrail
      I_Contact( "DI_INPUTS".R17_INPUTS_RUA.EMG_PB )
   END_RUNG wire#w4
   RUNG wire#powerrail
      Contact( "AlwaysTRUE" )
      wire#w5
      { S7_Templates := "SrcType := Int" } EQ_Contact(in1 := "Valves Data".R17_XV02.STATUS, in2 := 1)
      wire#w6
      Coil( "dummy".R17.Intl_1 )
   END_RUNG
   RUNG wire#w5
      { S7_Templates := "SrcType := Int" } EQ_Contact(in1 := "Valves Data".R17_XV03.STATUS, in2 := 1)
   END_RUNG wire#w6
   RUNG wire#w5
      { S7_Templates := "SrcType := Int" } EQ_Contact(in1 := "Valves Data".R17_XV04.STATUS, in2 := 1)
   END_RUNG wire#w6
   // the same network as SCL:
   IF "AlwaysTRUE" THEN
       #valve_R17_XV01("auto/manual" := "Valves Data"."A/M".R17,   // "valve"
                       open_auto := "R17_DATA".R17.HWS_CMD_2 OR "R17_DATA".R17.HWS_CMD_1,
                       open_man := "Valves Data".R17_XV01.MCMD AND NOT "dummy".R17.Intl_1,
                       fbk_open := "A/SSR_017_XV651_OFB",
                       fbk_close := "A/SSR_017_XV651_CFB",
                       reset := "Valves Data".R17_XV01.RESET OR "R17_DATA".R17.Reset,
                       intl := NOT "DI_INPUTS".R17_INPUTS_RUA.EMG_PB,
                       Mon_En := 1,
                       mon_sp := "Valves Data".R17_XV01.MON_TIME,
                       SEMI := "Valves Data".SEMI_AUTO.R17,
                       "open/close" => "A/SSR_017_XV651_CMD",
                       FAIL_TO_OPEN => "Valves Data".R17_VALVE_FAULT.XV01_FAIL_TO_OPEN,
                       FAIL_TO_CLOSE => "Valves Data".R17_VALVE_FAULT.XV01_FAIL_TO_CLOSE,
                       status => "Valves Data".R17_XV01.STATUS);
   END_IF;
   "dummy".R17.Intl_1 := "AlwaysTRUE" AND (("Valves Data".R17_XV02.STATUS = 1) OR ("Valves Data".R17_XV03.STATUS = 1) OR ("Valves Data".R17_XV04.STATUS = 1));
END_REGION

REGION Network 177: R17_XV02
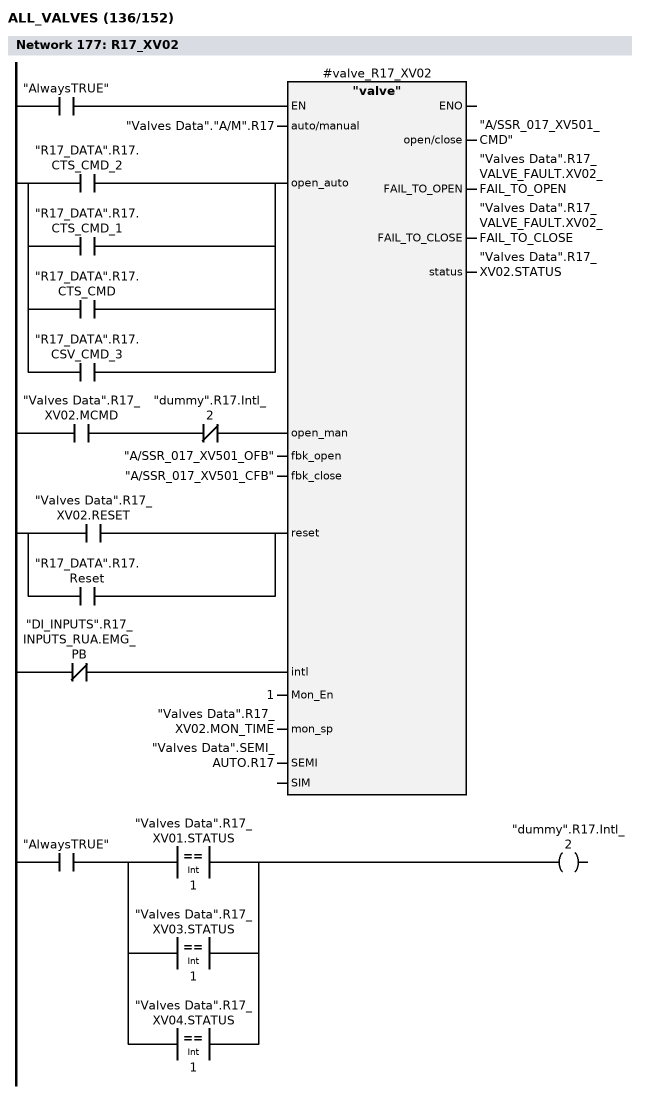
   RUNG wire#powerrail
      Contact( "AlwaysTRUE" )
      #valve_R17_XV02(open_auto := wire#w1, open_man := wire#w2, reset := wire#w3, intl := wire#w4, "auto/manual" := "Valves Data"."A/M".R17, fbk_open := "A/SSR_017_XV501_OFB", fbk_close := "A/SSR_017_XV501_CFB", Mon_En := 1, mon_sp := "Valves Data".R17_XV02.MON_TIME, SEMI := "Valves Data".SEMI_AUTO.R17, SIM :=, "open/close" => "A/SSR_017_XV501_CMD", FAIL_TO_OPEN => "Valves Data".R17_VALVE_FAULT.XV02_FAIL_TO_OPEN, FAIL_TO_CLOSE => "Valves Data".R17_VALVE_FAULT.XV02_FAIL_TO_CLOSE, status => "Valves Data".R17_XV02.STATUS)
   END_RUNG
   RUNG wire#powerrail
      Contact( "R17_DATA".R17.CTS_CMD_2 )
   END_RUNG wire#w1
   RUNG wire#powerrail
      Contact( "R17_DATA".R17.CTS_CMD_1 )
   END_RUNG wire#w1
   RUNG wire#powerrail
      Contact( "R17_DATA".R17.CTS_CMD )
   END_RUNG wire#w1
   RUNG wire#powerrail
      Contact( "R17_DATA".R17.CSV_CMD_3 )
   END_RUNG wire#w1
   RUNG wire#powerrail
      Contact( "Valves Data".R17_XV02.MCMD )
      I_Contact( "dummy".R17.Intl_2 )
   END_RUNG wire#w2
   RUNG wire#powerrail
      Contact( "Valves Data".R17_XV02.RESET )
   END_RUNG wire#w3
   RUNG wire#powerrail
      Contact( "R17_DATA".R17.Reset )
   END_RUNG wire#w3
   RUNG wire#powerrail
      I_Contact( "DI_INPUTS".R17_INPUTS_RUA.EMG_PB )
   END_RUNG wire#w4
   RUNG wire#powerrail
      Contact( "AlwaysTRUE" )
      wire#w5
      { S7_Templates := "SrcType := Int" } EQ_Contact(in1 := "Valves Data".R17_XV01.STATUS, in2 := 1)
      wire#w6
      Coil( "dummy".R17.Intl_2 )
   END_RUNG
   RUNG wire#w5
      { S7_Templates := "SrcType := Int" } EQ_Contact(in1 := "Valves Data".R17_XV03.STATUS, in2 := 1)
   END_RUNG wire#w6
   RUNG wire#w5
      { S7_Templates := "SrcType := Int" } EQ_Contact(in1 := "Valves Data".R17_XV04.STATUS, in2 := 1)
   END_RUNG wire#w6
   // the same network as SCL:
   IF "AlwaysTRUE" THEN
       #valve_R17_XV02("auto/manual" := "Valves Data"."A/M".R17,   // "valve"
                       open_auto := "R17_DATA".R17.CTS_CMD_2 OR "R17_DATA".R17.CTS_CMD_1 OR "R17_DATA".R17.CTS_CMD OR "R17_DATA".R17.CSV_CMD_3,
                       open_man := "Valves Data".R17_XV02.MCMD AND NOT "dummy".R17.Intl_2,
                       fbk_open := "A/SSR_017_XV501_OFB",
                       fbk_close := "A/SSR_017_XV501_CFB",
                       reset := "Valves Data".R17_XV02.RESET OR "R17_DATA".R17.Reset,
                       intl := NOT "DI_INPUTS".R17_INPUTS_RUA.EMG_PB,
                       Mon_En := 1,
                       mon_sp := "Valves Data".R17_XV02.MON_TIME,
                       SEMI := "Valves Data".SEMI_AUTO.R17,
                       "open/close" => "A/SSR_017_XV501_CMD",
                       FAIL_TO_OPEN => "Valves Data".R17_VALVE_FAULT.XV02_FAIL_TO_OPEN,
                       FAIL_TO_CLOSE => "Valves Data".R17_VALVE_FAULT.XV02_FAIL_TO_CLOSE,
                       status => "Valves Data".R17_XV02.STATUS);
   END_IF;
   "dummy".R17.Intl_2 := "AlwaysTRUE" AND (("Valves Data".R17_XV01.STATUS = 1) OR ("Valves Data".R17_XV03.STATUS = 1) OR ("Valves Data".R17_XV04.STATUS = 1));
END_REGION

REGION Network 178: R17_XV03
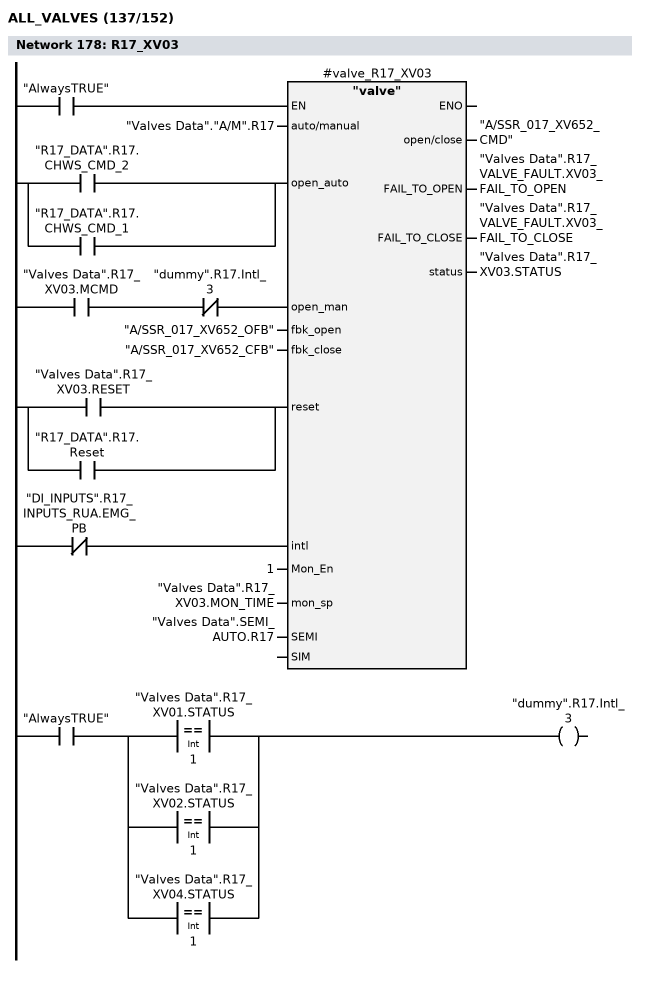
   RUNG wire#powerrail
      Contact( "AlwaysTRUE" )
      #valve_R17_XV03(open_auto := wire#w1, open_man := wire#w2, reset := wire#w3, intl := wire#w4, "auto/manual" := "Valves Data"."A/M".R17, fbk_open := "A/SSR_017_XV652_OFB", fbk_close := "A/SSR_017_XV652_CFB", Mon_En := 1, mon_sp := "Valves Data".R17_XV03.MON_TIME, SEMI := "Valves Data".SEMI_AUTO.R17, SIM :=, "open/close" => "A/SSR_017_XV652_CMD", FAIL_TO_OPEN => "Valves Data".R17_VALVE_FAULT.XV03_FAIL_TO_OPEN, FAIL_TO_CLOSE => "Valves Data".R17_VALVE_FAULT.XV03_FAIL_TO_CLOSE, status => "Valves Data".R17_XV03.STATUS)
   END_RUNG
   RUNG wire#powerrail
      Contact( "R17_DATA".R17.CHWS_CMD_2 )
   END_RUNG wire#w1
   RUNG wire#powerrail
      Contact( "R17_DATA".R17.CHWS_CMD_1 )
   END_RUNG wire#w1
   RUNG wire#powerrail
      Contact( "Valves Data".R17_XV03.MCMD )
      I_Contact( "dummy".R17.Intl_3 )
   END_RUNG wire#w2
   RUNG wire#powerrail
      Contact( "Valves Data".R17_XV03.RESET )
   END_RUNG wire#w3
   RUNG wire#powerrail
      Contact( "R17_DATA".R17.Reset )
   END_RUNG wire#w3
   RUNG wire#powerrail
      I_Contact( "DI_INPUTS".R17_INPUTS_RUA.EMG_PB )
   END_RUNG wire#w4
   RUNG wire#powerrail
      Contact( "AlwaysTRUE" )
      wire#w5
      { S7_Templates := "SrcType := Int" } EQ_Contact(in1 := "Valves Data".R17_XV01.STATUS, in2 := 1)
      wire#w6
      Coil( "dummy".R17.Intl_3 )
   END_RUNG
   RUNG wire#w5
      { S7_Templates := "SrcType := Int" } EQ_Contact(in1 := "Valves Data".R17_XV02.STATUS, in2 := 1)
   END_RUNG wire#w6
   RUNG wire#w5
      { S7_Templates := "SrcType := Int" } EQ_Contact(in1 := "Valves Data".R17_XV04.STATUS, in2 := 1)
   END_RUNG wire#w6
   // the same network as SCL:
   IF "AlwaysTRUE" THEN
       #valve_R17_XV03("auto/manual" := "Valves Data"."A/M".R17,   // "valve"
                       open_auto := "R17_DATA".R17.CHWS_CMD_2 OR "R17_DATA".R17.CHWS_CMD_1,
                       open_man := "Valves Data".R17_XV03.MCMD AND NOT "dummy".R17.Intl_3,
                       fbk_open := "A/SSR_017_XV652_OFB",
                       fbk_close := "A/SSR_017_XV652_CFB",
                       reset := "Valves Data".R17_XV03.RESET OR "R17_DATA".R17.Reset,
                       intl := NOT "DI_INPUTS".R17_INPUTS_RUA.EMG_PB,
                       Mon_En := 1,
                       mon_sp := "Valves Data".R17_XV03.MON_TIME,
                       SEMI := "Valves Data".SEMI_AUTO.R17,
                       "open/close" => "A/SSR_017_XV652_CMD",
                       FAIL_TO_OPEN => "Valves Data".R17_VALVE_FAULT.XV03_FAIL_TO_OPEN,
                       FAIL_TO_CLOSE => "Valves Data".R17_VALVE_FAULT.XV03_FAIL_TO_CLOSE,
                       status => "Valves Data".R17_XV03.STATUS);
   END_IF;
   "dummy".R17.Intl_3 := "AlwaysTRUE" AND (("Valves Data".R17_XV01.STATUS = 1) OR ("Valves Data".R17_XV02.STATUS = 1) OR ("Valves Data".R17_XV04.STATUS = 1));
END_REGION

REGION Network 179: R17_XV04
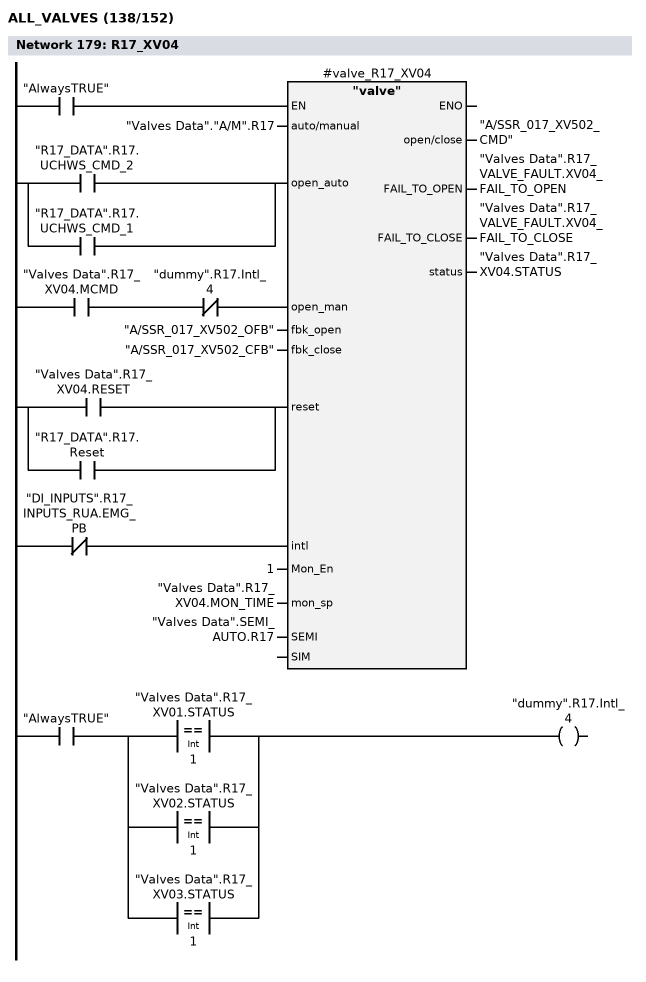
   RUNG wire#powerrail
      Contact( "AlwaysTRUE" )
      #valve_R17_XV04(open_auto := wire#w1, open_man := wire#w2, reset := wire#w3, intl := wire#w4, "auto/manual" := "Valves Data"."A/M".R17, fbk_open := "A/SSR_017_XV502_OFB", fbk_close := "A/SSR_017_XV502_CFB", Mon_En := 1, mon_sp := "Valves Data".R17_XV04.MON_TIME, SEMI := "Valves Data".SEMI_AUTO.R17, SIM :=, "open/close" => "A/SSR_017_XV502_CMD", FAIL_TO_OPEN => "Valves Data".R17_VALVE_FAULT.XV04_FAIL_TO_OPEN, FAIL_TO_CLOSE => "Valves Data".R17_VALVE_FAULT.XV04_FAIL_TO_CLOSE, status => "Valves Data".R17_XV04.STATUS)
   END_RUNG
   RUNG wire#powerrail
      Contact( "R17_DATA".R17.UCHWS_CMD_2 )
   END_RUNG wire#w1
   RUNG wire#powerrail
      Contact( "R17_DATA".R17.UCHWS_CMD_1 )
   END_RUNG wire#w1
   RUNG wire#powerrail
      Contact( "Valves Data".R17_XV04.MCMD )
      I_Contact( "dummy".R17.Intl_4 )
   END_RUNG wire#w2
   RUNG wire#powerrail
      Contact( "Valves Data".R17_XV04.RESET )
   END_RUNG wire#w3
   RUNG wire#powerrail
      Contact( "R17_DATA".R17.Reset )
   END_RUNG wire#w3
   RUNG wire#powerrail
      I_Contact( "DI_INPUTS".R17_INPUTS_RUA.EMG_PB )
   END_RUNG wire#w4
   RUNG wire#powerrail
      Contact( "AlwaysTRUE" )
      wire#w5
      { S7_Templates := "SrcType := Int" } EQ_Contact(in1 := "Valves Data".R17_XV01.STATUS, in2 := 1)
      wire#w6
      Coil( "dummy".R17.Intl_4 )
   END_RUNG
   RUNG wire#w5
      { S7_Templates := "SrcType := Int" } EQ_Contact(in1 := "Valves Data".R17_XV02.STATUS, in2 := 1)
   END_RUNG wire#w6
   RUNG wire#w5
      { S7_Templates := "SrcType := Int" } EQ_Contact(in1 := "Valves Data".R17_XV03.STATUS, in2 := 1)
   END_RUNG wire#w6
   // the same network as SCL:
   IF "AlwaysTRUE" THEN
       #valve_R17_XV04("auto/manual" := "Valves Data"."A/M".R17,   // "valve"
                       open_auto := "R17_DATA".R17.UCHWS_CMD_2 OR "R17_DATA".R17.UCHWS_CMD_1,
                       open_man := "Valves Data".R17_XV04.MCMD AND NOT "dummy".R17.Intl_4,
                       fbk_open := "A/SSR_017_XV502_OFB",
                       fbk_close := "A/SSR_017_XV502_CFB",
                       reset := "Valves Data".R17_XV04.RESET OR "R17_DATA".R17.Reset,
                       intl := NOT "DI_INPUTS".R17_INPUTS_RUA.EMG_PB,
                       Mon_En := 1,
                       mon_sp := "Valves Data".R17_XV04.MON_TIME,
                       SEMI := "Valves Data".SEMI_AUTO.R17,
                       "open/close" => "A/SSR_017_XV502_CMD",
                       FAIL_TO_OPEN => "Valves Data".R17_VALVE_FAULT.XV04_FAIL_TO_OPEN,
                       FAIL_TO_CLOSE => "Valves Data".R17_VALVE_FAULT.XV04_FAIL_TO_CLOSE,
                       status => "Valves Data".R17_XV04.STATUS);
   END_IF;
   "dummy".R17.Intl_4 := "AlwaysTRUE" AND (("Valves Data".R17_XV01.STATUS = 1) OR ("Valves Data".R17_XV02.STATUS = 1) OR ("Valves Data".R17_XV03.STATUS = 1));
END_REGION

REGION Network 180: R17_XV05
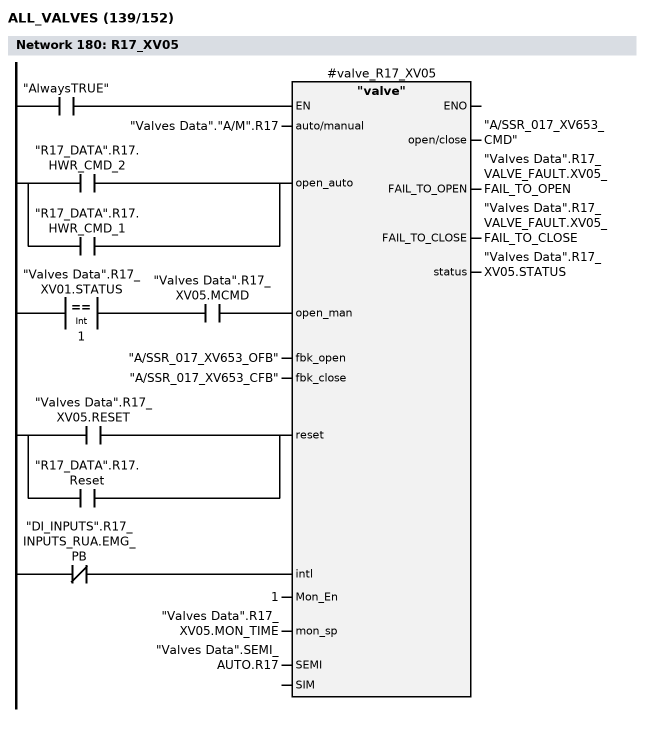
   RUNG wire#powerrail
      Contact( "AlwaysTRUE" )
      #valve_R17_XV05(open_auto := wire#w1, open_man := wire#w2, reset := wire#w3, intl := wire#w4, "auto/manual" := "Valves Data"."A/M".R17, fbk_open := "A/SSR_017_XV653_OFB", fbk_close := "A/SSR_017_XV653_CFB", Mon_En := 1, mon_sp := "Valves Data".R17_XV05.MON_TIME, SEMI := "Valves Data".SEMI_AUTO.R17, SIM :=, "open/close" => "A/SSR_017_XV653_CMD", FAIL_TO_OPEN => "Valves Data".R17_VALVE_FAULT.XV05_FAIL_TO_OPEN, FAIL_TO_CLOSE => "Valves Data".R17_VALVE_FAULT.XV05_FAIL_TO_CLOSE, status => "Valves Data".R17_XV05.STATUS)
   END_RUNG
   RUNG wire#powerrail
      Contact( "R17_DATA".R17.HWR_CMD_2 )
   END_RUNG wire#w1
   RUNG wire#powerrail
      Contact( "R17_DATA".R17.HWR_CMD_1 )
   END_RUNG wire#w1
   RUNG wire#powerrail
      { S7_Templates := "SrcType := Int" } EQ_Contact(in1 := "Valves Data".R17_XV01.STATUS, in2 := 1)
      Contact( "Valves Data".R17_XV05.MCMD )
   END_RUNG wire#w2
   RUNG wire#powerrail
      Contact( "Valves Data".R17_XV05.RESET )
   END_RUNG wire#w3
   RUNG wire#powerrail
      Contact( "R17_DATA".R17.Reset )
   END_RUNG wire#w3
   RUNG wire#powerrail
      I_Contact( "DI_INPUTS".R17_INPUTS_RUA.EMG_PB )
   END_RUNG wire#w4
   // the same network as SCL:
   IF "AlwaysTRUE" THEN
       #valve_R17_XV05("auto/manual" := "Valves Data"."A/M".R17,   // "valve"
                       open_auto := "R17_DATA".R17.HWR_CMD_2 OR "R17_DATA".R17.HWR_CMD_1,
                       open_man := ("Valves Data".R17_XV01.STATUS = 1) AND "Valves Data".R17_XV05.MCMD,
                       fbk_open := "A/SSR_017_XV653_OFB",
                       fbk_close := "A/SSR_017_XV653_CFB",
                       reset := "Valves Data".R17_XV05.RESET OR "R17_DATA".R17.Reset,
                       intl := NOT "DI_INPUTS".R17_INPUTS_RUA.EMG_PB,
                       Mon_En := 1,
                       mon_sp := "Valves Data".R17_XV05.MON_TIME,
                       SEMI := "Valves Data".SEMI_AUTO.R17,
                       "open/close" => "A/SSR_017_XV653_CMD",
                       FAIL_TO_OPEN => "Valves Data".R17_VALVE_FAULT.XV05_FAIL_TO_OPEN,
                       FAIL_TO_CLOSE => "Valves Data".R17_VALVE_FAULT.XV05_FAIL_TO_CLOSE,
                       status => "Valves Data".R17_XV05.STATUS);
   END_IF;
END_REGION

REGION Network 181: R17_XV06
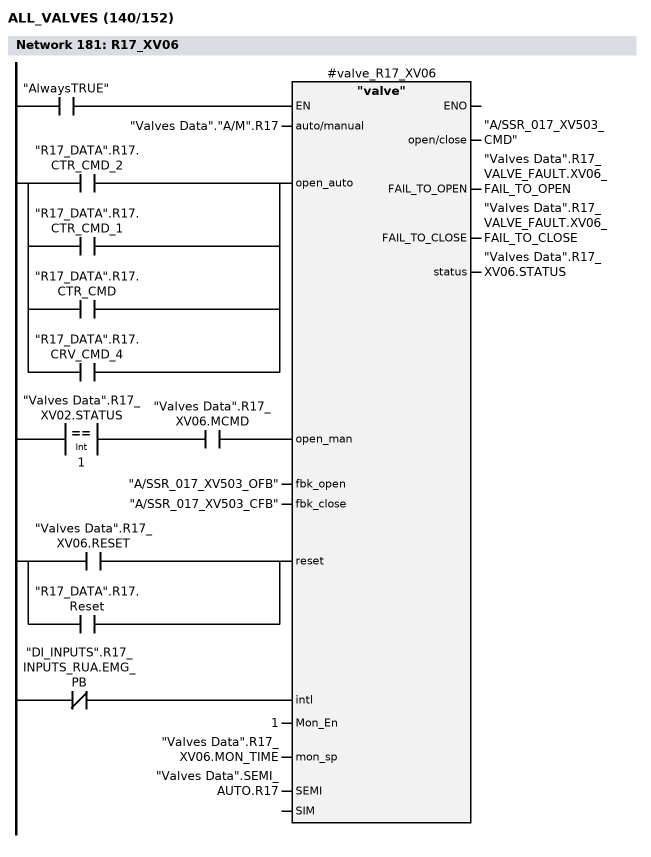
   RUNG wire#powerrail
      Contact( "AlwaysTRUE" )
      #valve_R17_XV06(open_auto := wire#w1, open_man := wire#w2, reset := wire#w3, intl := wire#w4, "auto/manual" := "Valves Data"."A/M".R17, fbk_open := "A/SSR_017_XV503_OFB", fbk_close := "A/SSR_017_XV503_CFB", Mon_En := 1, mon_sp := "Valves Data".R17_XV06.MON_TIME, SEMI := "Valves Data".SEMI_AUTO.R17, SIM :=, "open/close" => "A/SSR_017_XV503_CMD", FAIL_TO_OPEN => "Valves Data".R17_VALVE_FAULT.XV06_FAIL_TO_OPEN, FAIL_TO_CLOSE => "Valves Data".R17_VALVE_FAULT.XV06_FAIL_TO_CLOSE, status => "Valves Data".R17_XV06.STATUS)
   END_RUNG
   RUNG wire#powerrail
      Contact( "R17_DATA".R17.CTR_CMD_2 )
   END_RUNG wire#w1
   RUNG wire#powerrail
      Contact( "R17_DATA".R17.CTR_CMD_1 )
   END_RUNG wire#w1
   RUNG wire#powerrail
      Contact( "R17_DATA".R17.CTR_CMD )
   END_RUNG wire#w1
   RUNG wire#powerrail
      Contact( "R17_DATA".R17.CRV_CMD_4 )
   END_RUNG wire#w1
   RUNG wire#powerrail
      { S7_Templates := "SrcType := Int" } EQ_Contact(in1 := "Valves Data".R17_XV02.STATUS, in2 := 1)
      Contact( "Valves Data".R17_XV06.MCMD )
   END_RUNG wire#w2
   RUNG wire#powerrail
      Contact( "Valves Data".R17_XV06.RESET )
   END_RUNG wire#w3
   RUNG wire#powerrail
      Contact( "R17_DATA".R17.Reset )
   END_RUNG wire#w3
   RUNG wire#powerrail
      I_Contact( "DI_INPUTS".R17_INPUTS_RUA.EMG_PB )
   END_RUNG wire#w4
   // the same network as SCL:
   IF "AlwaysTRUE" THEN
       #valve_R17_XV06("auto/manual" := "Valves Data"."A/M".R17,   // "valve"
                       open_auto := "R17_DATA".R17.CTR_CMD_2 OR "R17_DATA".R17.CTR_CMD_1 OR "R17_DATA".R17.CTR_CMD OR "R17_DATA".R17.CRV_CMD_4,
                       open_man := ("Valves Data".R17_XV02.STATUS = 1) AND "Valves Data".R17_XV06.MCMD,
                       fbk_open := "A/SSR_017_XV503_OFB",
                       fbk_close := "A/SSR_017_XV503_CFB",
                       reset := "Valves Data".R17_XV06.RESET OR "R17_DATA".R17.Reset,
                       intl := NOT "DI_INPUTS".R17_INPUTS_RUA.EMG_PB,
                       Mon_En := 1,
                       mon_sp := "Valves Data".R17_XV06.MON_TIME,
                       SEMI := "Valves Data".SEMI_AUTO.R17,
                       "open/close" => "A/SSR_017_XV503_CMD",
                       FAIL_TO_OPEN => "Valves Data".R17_VALVE_FAULT.XV06_FAIL_TO_OPEN,
                       FAIL_TO_CLOSE => "Valves Data".R17_VALVE_FAULT.XV06_FAIL_TO_CLOSE,
                       status => "Valves Data".R17_XV06.STATUS);
   END_IF;
END_REGION

REGION Network 182: R17_XV07
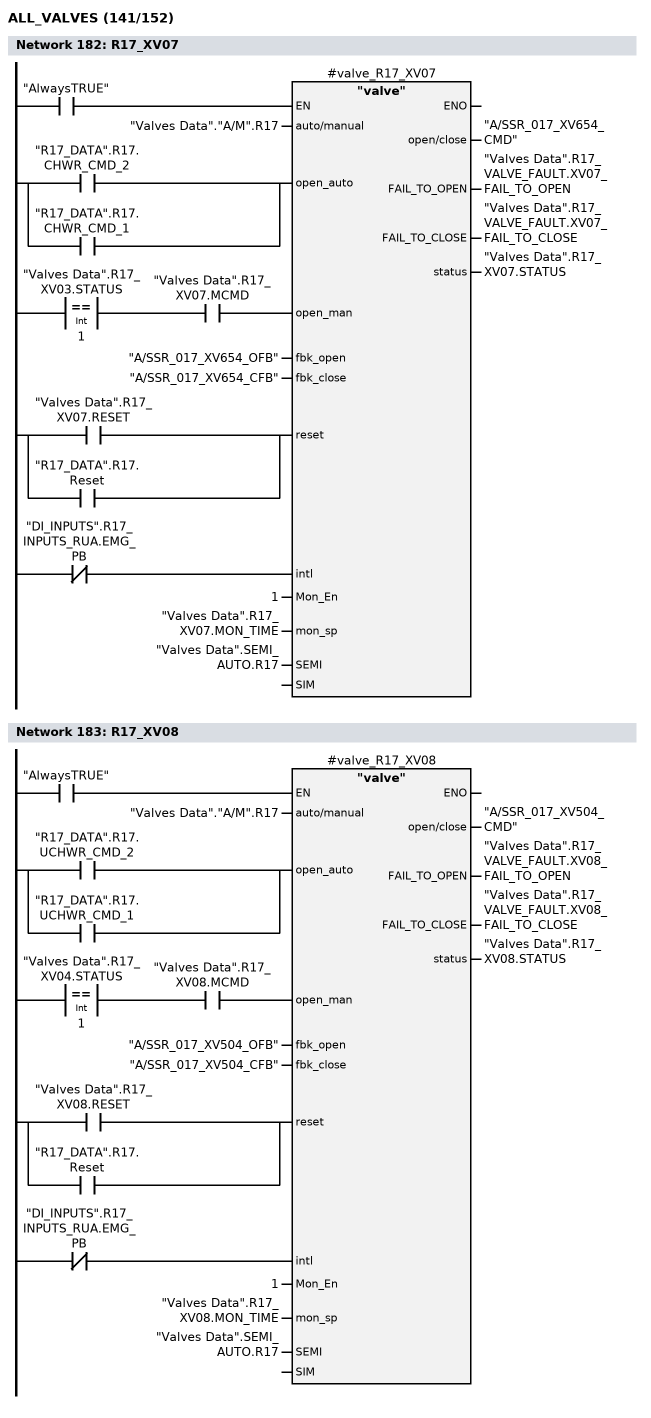
   RUNG wire#powerrail
      Contact( "AlwaysTRUE" )
      #valve_R17_XV07(open_auto := wire#w1, open_man := wire#w2, reset := wire#w3, intl := wire#w4, "auto/manual" := "Valves Data"."A/M".R17, fbk_open := "A/SSR_017_XV654_OFB", fbk_close := "A/SSR_017_XV654_CFB", Mon_En := 1, mon_sp := "Valves Data".R17_XV07.MON_TIME, SEMI := "Valves Data".SEMI_AUTO.R17, SIM :=, "open/close" => "A/SSR_017_XV654_CMD", FAIL_TO_OPEN => "Valves Data".R17_VALVE_FAULT.XV07_FAIL_TO_OPEN, FAIL_TO_CLOSE => "Valves Data".R17_VALVE_FAULT.XV07_FAIL_TO_CLOSE, status => "Valves Data".R17_XV07.STATUS)
   END_RUNG
   RUNG wire#powerrail
      Contact( "R17_DATA".R17.CHWR_CMD_2 )
   END_RUNG wire#w1
   RUNG wire#powerrail
      Contact( "R17_DATA".R17.CHWR_CMD_1 )
   END_RUNG wire#w1
   RUNG wire#powerrail
      { S7_Templates := "SrcType := Int" } EQ_Contact(in1 := "Valves Data".R17_XV03.STATUS, in2 := 1)
      Contact( "Valves Data".R17_XV07.MCMD )
   END_RUNG wire#w2
   RUNG wire#powerrail
      Contact( "Valves Data".R17_XV07.RESET )
   END_RUNG wire#w3
   RUNG wire#powerrail
      Contact( "R17_DATA".R17.Reset )
   END_RUNG wire#w3
   RUNG wire#powerrail
      I_Contact( "DI_INPUTS".R17_INPUTS_RUA.EMG_PB )
   END_RUNG wire#w4
   // the same network as SCL:
   IF "AlwaysTRUE" THEN
       #valve_R17_XV07("auto/manual" := "Valves Data"."A/M".R17,   // "valve"
                       open_auto := "R17_DATA".R17.CHWR_CMD_2 OR "R17_DATA".R17.CHWR_CMD_1,
                       open_man := ("Valves Data".R17_XV03.STATUS = 1) AND "Valves Data".R17_XV07.MCMD,
                       fbk_open := "A/SSR_017_XV654_OFB",
                       fbk_close := "A/SSR_017_XV654_CFB",
                       reset := "Valves Data".R17_XV07.RESET OR "R17_DATA".R17.Reset,
                       intl := NOT "DI_INPUTS".R17_INPUTS_RUA.EMG_PB,
                       Mon_En := 1,
                       mon_sp := "Valves Data".R17_XV07.MON_TIME,
                       SEMI := "Valves Data".SEMI_AUTO.R17,
                       "open/close" => "A/SSR_017_XV654_CMD",
                       FAIL_TO_OPEN => "Valves Data".R17_VALVE_FAULT.XV07_FAIL_TO_OPEN,
                       FAIL_TO_CLOSE => "Valves Data".R17_VALVE_FAULT.XV07_FAIL_TO_CLOSE,
                       status => "Valves Data".R17_XV07.STATUS);
   END_IF;
END_REGION

REGION Network 183: R17_XV08
   RUNG wire#powerrail
      Contact( "AlwaysTRUE" )
      #valve_R17_XV08(open_auto := wire#w1, open_man := wire#w2, reset := wire#w3, intl := wire#w4, "auto/manual" := "Valves Data"."A/M".R17, fbk_open := "A/SSR_017_XV504_OFB", fbk_close := "A/SSR_017_XV504_CFB", Mon_En := 1, mon_sp := "Valves Data".R17_XV08.MON_TIME, SEMI := "Valves Data".SEMI_AUTO.R17, SIM :=, "open/close" => "A/SSR_017_XV504_CMD", FAIL_TO_OPEN => "Valves Data".R17_VALVE_FAULT.XV08_FAIL_TO_OPEN, FAIL_TO_CLOSE => "Valves Data".R17_VALVE_FAULT.XV08_FAIL_TO_CLOSE, status => "Valves Data".R17_XV08.STATUS)
   END_RUNG
   RUNG wire#powerrail
      Contact( "R17_DATA".R17.UCHWR_CMD_2 )
   END_RUNG wire#w1
   RUNG wire#powerrail
      Contact( "R17_DATA".R17.UCHWR_CMD_1 )
   END_RUNG wire#w1
   RUNG wire#powerrail
      { S7_Templates := "SrcType := Int" } EQ_Contact(in1 := "Valves Data".R17_XV04.STATUS, in2 := 1)
      Contact( "Valves Data".R17_XV08.MCMD )
   END_RUNG wire#w2
   RUNG wire#powerrail
      Contact( "Valves Data".R17_XV08.RESET )
   END_RUNG wire#w3
   RUNG wire#powerrail
      Contact( "R17_DATA".R17.Reset )
   END_RUNG wire#w3
   RUNG wire#powerrail
      I_Contact( "DI_INPUTS".R17_INPUTS_RUA.EMG_PB )
   END_RUNG wire#w4
   // the same network as SCL:
   IF "AlwaysTRUE" THEN
       #valve_R17_XV08("auto/manual" := "Valves Data"."A/M".R17,   // "valve"
                       open_auto := "R17_DATA".R17.UCHWR_CMD_2 OR "R17_DATA".R17.UCHWR_CMD_1,
                       open_man := ("Valves Data".R17_XV04.STATUS = 1) AND "Valves Data".R17_XV08.MCMD,
                       fbk_open := "A/SSR_017_XV504_OFB",
                       fbk_close := "A/SSR_017_XV504_CFB",
                       reset := "Valves Data".R17_XV08.RESET OR "R17_DATA".R17.Reset,
                       intl := NOT "DI_INPUTS".R17_INPUTS_RUA.EMG_PB,
                       Mon_En := 1,
                       mon_sp := "Valves Data".R17_XV08.MON_TIME,
                       SEMI := "Valves Data".SEMI_AUTO.R17,
                       "open/close" => "A/SSR_017_XV504_CMD",
                       FAIL_TO_OPEN => "Valves Data".R17_VALVE_FAULT.XV08_FAIL_TO_OPEN,
                       FAIL_TO_CLOSE => "Valves Data".R17_VALVE_FAULT.XV08_FAIL_TO_CLOSE,
                       status => "Valves Data".R17_XV08.STATUS);
   END_IF;
END_REGION

REGION Network 184: R17_XV09
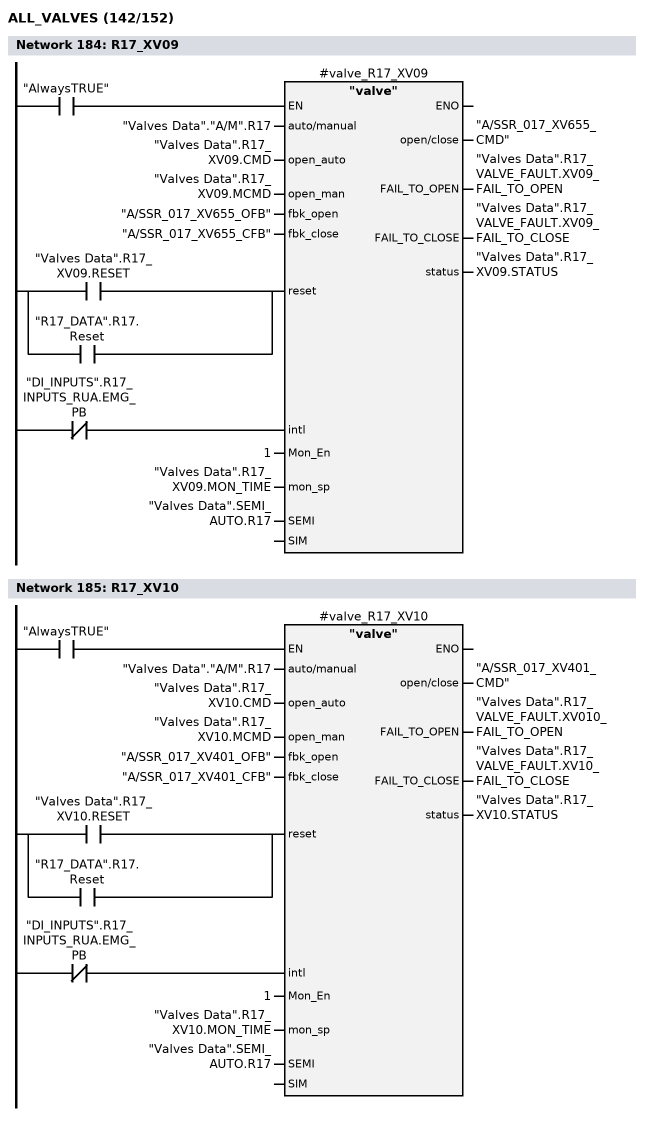
   RUNG wire#powerrail
      Contact( "AlwaysTRUE" )
      #valve_R17_XV09(reset := wire#w1, intl := wire#w2, "auto/manual" := "Valves Data"."A/M".R17, open_auto := "Valves Data".R17_XV09.CMD, open_man := "Valves Data".R17_XV09.MCMD, fbk_open := "A/SSR_017_XV655_OFB", fbk_close := "A/SSR_017_XV655_CFB", Mon_En := 1, mon_sp := "Valves Data".R17_XV09.MON_TIME, SEMI := "Valves Data".SEMI_AUTO.R17, SIM :=, "open/close" => "A/SSR_017_XV655_CMD", FAIL_TO_OPEN => "Valves Data".R17_VALVE_FAULT.XV09_FAIL_TO_OPEN, FAIL_TO_CLOSE => "Valves Data".R17_VALVE_FAULT.XV09_FAIL_TO_CLOSE, status => "Valves Data".R17_XV09.STATUS)
   END_RUNG
   RUNG wire#powerrail
      Contact( "Valves Data".R17_XV09.RESET )
   END_RUNG wire#w1
   RUNG wire#powerrail
      Contact( "R17_DATA".R17.Reset )
   END_RUNG wire#w1
   RUNG wire#powerrail
      I_Contact( "DI_INPUTS".R17_INPUTS_RUA.EMG_PB )
   END_RUNG wire#w2
   // the same network as SCL:
   IF "AlwaysTRUE" THEN
       #valve_R17_XV09("auto/manual" := "Valves Data"."A/M".R17,   // "valve"
                       open_auto := "Valves Data".R17_XV09.CMD,
                       open_man := "Valves Data".R17_XV09.MCMD,
                       fbk_open := "A/SSR_017_XV655_OFB",
                       fbk_close := "A/SSR_017_XV655_CFB",
                       reset := "Valves Data".R17_XV09.RESET OR "R17_DATA".R17.Reset,
                       intl := NOT "DI_INPUTS".R17_INPUTS_RUA.EMG_PB,
                       Mon_En := 1,
                       mon_sp := "Valves Data".R17_XV09.MON_TIME,
                       SEMI := "Valves Data".SEMI_AUTO.R17,
                       "open/close" => "A/SSR_017_XV655_CMD",
                       FAIL_TO_OPEN => "Valves Data".R17_VALVE_FAULT.XV09_FAIL_TO_OPEN,
                       FAIL_TO_CLOSE => "Valves Data".R17_VALVE_FAULT.XV09_FAIL_TO_CLOSE,
                       status => "Valves Data".R17_XV09.STATUS);
   END_IF;
END_REGION

REGION Network 185: R17_XV10
   RUNG wire#powerrail
      Contact( "AlwaysTRUE" )
      #valve_R17_XV10(reset := wire#w1, intl := wire#w2, "auto/manual" := "Valves Data"."A/M".R17, open_auto := "Valves Data".R17_XV10.CMD, open_man := "Valves Data".R17_XV10.MCMD, fbk_open := "A/SSR_017_XV401_OFB", fbk_close := "A/SSR_017_XV401_CFB", Mon_En := 1, mon_sp := "Valves Data".R17_XV10.MON_TIME, SEMI := "Valves Data".SEMI_AUTO.R17, SIM :=, "open/close" => "A/SSR_017_XV401_CMD", FAIL_TO_OPEN => "Valves Data".R17_VALVE_FAULT.XV010_FAIL_TO_OPEN, FAIL_TO_CLOSE => "Valves Data".R17_VALVE_FAULT.XV10_FAIL_TO_CLOSE, status => "Valves Data".R17_XV10.STATUS)
   END_RUNG
   RUNG wire#powerrail
      Contact( "Valves Data".R17_XV10.RESET )
   END_RUNG wire#w1
   RUNG wire#powerrail
      Contact( "R17_DATA".R17.Reset )
   END_RUNG wire#w1
   RUNG wire#powerrail
      I_Contact( "DI_INPUTS".R17_INPUTS_RUA.EMG_PB )
   END_RUNG wire#w2
   // the same network as SCL:
   IF "AlwaysTRUE" THEN
       #valve_R17_XV10("auto/manual" := "Valves Data"."A/M".R17,   // "valve"
                       open_auto := "Valves Data".R17_XV10.CMD,
                       open_man := "Valves Data".R17_XV10.MCMD,
                       fbk_open := "A/SSR_017_XV401_OFB",
                       fbk_close := "A/SSR_017_XV401_CFB",
                       reset := "Valves Data".R17_XV10.RESET OR "R17_DATA".R17.Reset,
                       intl := NOT "DI_INPUTS".R17_INPUTS_RUA.EMG_PB,
                       Mon_En := 1,
                       mon_sp := "Valves Data".R17_XV10.MON_TIME,
                       SEMI := "Valves Data".SEMI_AUTO.R17,
                       "open/close" => "A/SSR_017_XV401_CMD",
                       FAIL_TO_OPEN => "Valves Data".R17_VALVE_FAULT.XV010_FAIL_TO_OPEN,
                       FAIL_TO_CLOSE => "Valves Data".R17_VALVE_FAULT.XV10_FAIL_TO_CLOSE,
                       status => "Valves Data".R17_XV10.STATUS);
   END_IF;
END_REGION

REGION Network 186: ****REACTOR_18****
END_REGION

REGION Network 187: R18_XV01
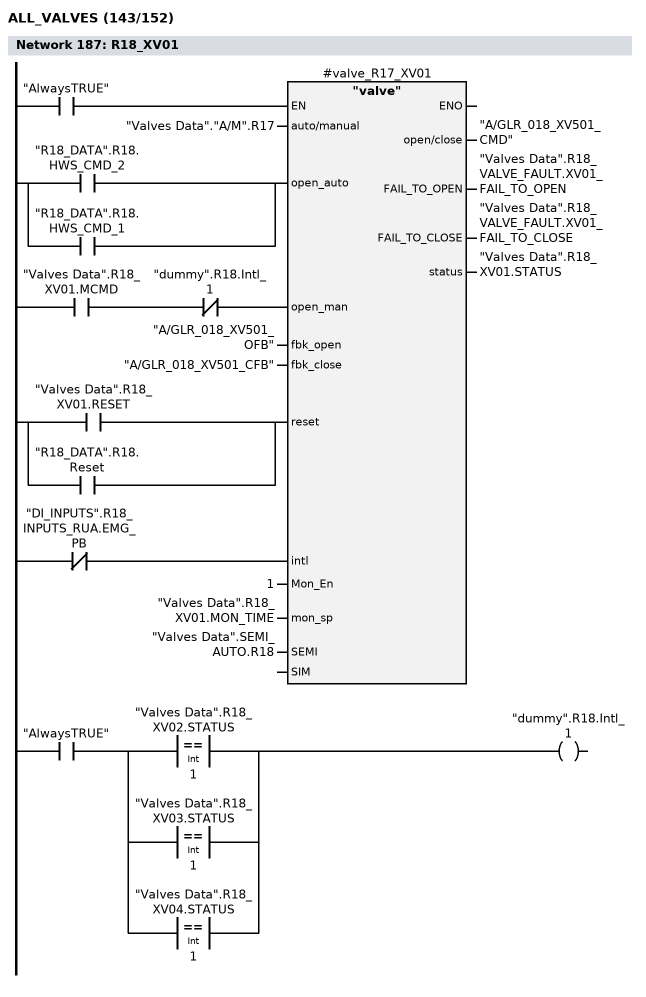
   RUNG wire#powerrail
      Contact( "AlwaysTRUE" )
      #valve_R17_XV01(open_auto := wire#w1, open_man := wire#w2, reset := wire#w3, intl := wire#w4, "auto/manual" := "Valves Data"."A/M".R17, fbk_open := "A/GLR_018_XV501_OFB", fbk_close := "A/GLR_018_XV501_CFB", Mon_En := 1, mon_sp := "Valves Data".R18_XV01.MON_TIME, SEMI := "Valves Data".SEMI_AUTO.R18, SIM :=, "open/close" => "A/GLR_018_XV501_CMD", FAIL_TO_OPEN => "Valves Data".R18_VALVE_FAULT.XV01_FAIL_TO_OPEN, FAIL_TO_CLOSE => "Valves Data".R18_VALVE_FAULT.XV01_FAIL_TO_CLOSE, status => "Valves Data".R18_XV01.STATUS)
   END_RUNG
   RUNG wire#powerrail
      Contact( "R18_DATA".R18.HWS_CMD_2 )
   END_RUNG wire#w1
   RUNG wire#powerrail
      Contact( "R18_DATA".R18.HWS_CMD_1 )
   END_RUNG wire#w1
   RUNG wire#powerrail
      Contact( "Valves Data".R18_XV01.MCMD )
      I_Contact( "dummy".R18.Intl_1 )
   END_RUNG wire#w2
   RUNG wire#powerrail
      Contact( "Valves Data".R18_XV01.RESET )
   END_RUNG wire#w3
   RUNG wire#powerrail
      Contact( "R18_DATA".R18.Reset )
   END_RUNG wire#w3
   RUNG wire#powerrail
      I_Contact( "DI_INPUTS".R18_INPUTS_RUA.EMG_PB )
   END_RUNG wire#w4
   RUNG wire#powerrail
      Contact( "AlwaysTRUE" )
      wire#w5
      { S7_Templates := "SrcType := Int" } EQ_Contact(in1 := "Valves Data".R18_XV02.STATUS, in2 := 1)
      wire#w6
      Coil( "dummy".R18.Intl_1 )
   END_RUNG
   RUNG wire#w5
      { S7_Templates := "SrcType := Int" } EQ_Contact(in1 := "Valves Data".R18_XV03.STATUS, in2 := 1)
   END_RUNG wire#w6
   RUNG wire#w5
      { S7_Templates := "SrcType := Int" } EQ_Contact(in1 := "Valves Data".R18_XV04.STATUS, in2 := 1)
   END_RUNG wire#w6
   // the same network as SCL:
   IF "AlwaysTRUE" THEN
       #valve_R17_XV01("auto/manual" := "Valves Data"."A/M".R17,   // "valve"
                       open_auto := "R18_DATA".R18.HWS_CMD_2 OR "R18_DATA".R18.HWS_CMD_1,
                       open_man := "Valves Data".R18_XV01.MCMD AND NOT "dummy".R18.Intl_1,
                       fbk_open := "A/GLR_018_XV501_OFB",
                       fbk_close := "A/GLR_018_XV501_CFB",
                       reset := "Valves Data".R18_XV01.RESET OR "R18_DATA".R18.Reset,
                       intl := NOT "DI_INPUTS".R18_INPUTS_RUA.EMG_PB,
                       Mon_En := 1,
                       mon_sp := "Valves Data".R18_XV01.MON_TIME,
                       SEMI := "Valves Data".SEMI_AUTO.R18,
                       "open/close" => "A/GLR_018_XV501_CMD",
                       FAIL_TO_OPEN => "Valves Data".R18_VALVE_FAULT.XV01_FAIL_TO_OPEN,
                       FAIL_TO_CLOSE => "Valves Data".R18_VALVE_FAULT.XV01_FAIL_TO_CLOSE,
                       status => "Valves Data".R18_XV01.STATUS);
   END_IF;
   "dummy".R18.Intl_1 := "AlwaysTRUE" AND (("Valves Data".R18_XV02.STATUS = 1) OR ("Valves Data".R18_XV03.STATUS = 1) OR ("Valves Data".R18_XV04.STATUS = 1));
END_REGION

REGION Network 188: R18_XV02
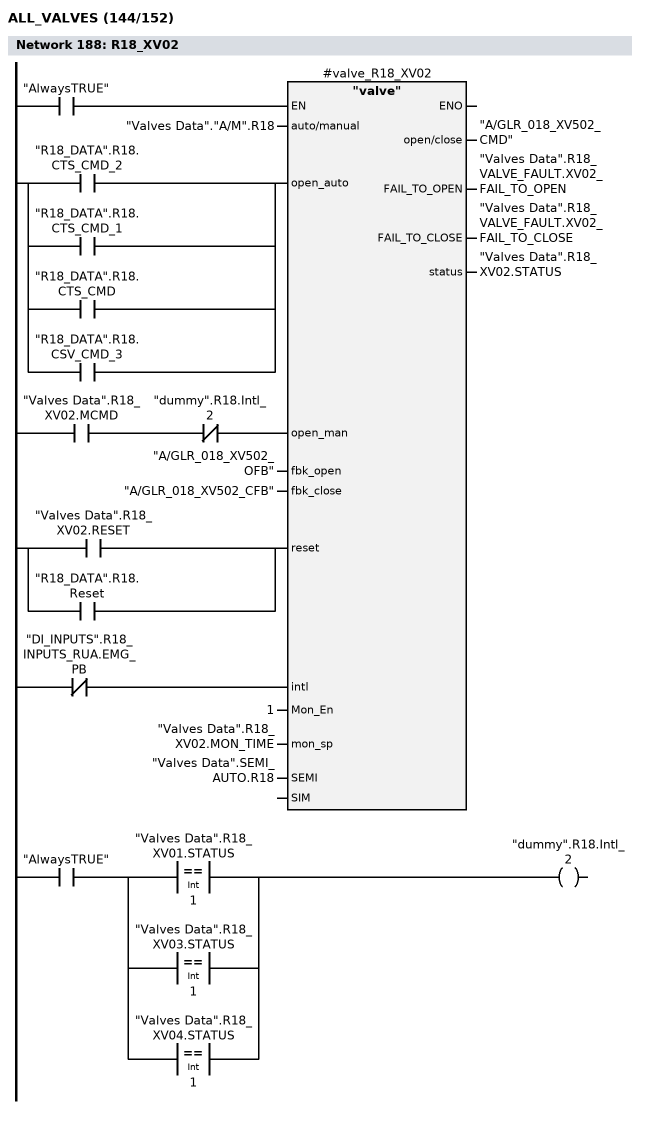
   RUNG wire#powerrail
      Contact( "AlwaysTRUE" )
      #valve_R18_XV02(open_auto := wire#w1, open_man := wire#w2, reset := wire#w3, intl := wire#w4, "auto/manual" := "Valves Data"."A/M".R18, fbk_open := "A/GLR_018_XV502_OFB", fbk_close := "A/GLR_018_XV502_CFB", Mon_En := 1, mon_sp := "Valves Data".R18_XV02.MON_TIME, SEMI := "Valves Data".SEMI_AUTO.R18, SIM :=, "open/close" => "A/GLR_018_XV502_CMD", FAIL_TO_OPEN => "Valves Data".R18_VALVE_FAULT.XV02_FAIL_TO_OPEN, FAIL_TO_CLOSE => "Valves Data".R18_VALVE_FAULT.XV02_FAIL_TO_CLOSE, status => "Valves Data".R18_XV02.STATUS)
   END_RUNG
   RUNG wire#powerrail
      Contact( "R18_DATA".R18.CTS_CMD_2 )
   END_RUNG wire#w1
   RUNG wire#powerrail
      Contact( "R18_DATA".R18.CTS_CMD_1 )
   END_RUNG wire#w1
   RUNG wire#powerrail
      Contact( "R18_DATA".R18.CTS_CMD )
   END_RUNG wire#w1
   RUNG wire#powerrail
      Contact( "R18_DATA".R18.CSV_CMD_3 )
   END_RUNG wire#w1
   RUNG wire#powerrail
      Contact( "Valves Data".R18_XV02.MCMD )
      I_Contact( "dummy".R18.Intl_2 )
   END_RUNG wire#w2
   RUNG wire#powerrail
      Contact( "Valves Data".R18_XV02.RESET )
   END_RUNG wire#w3
   RUNG wire#powerrail
      Contact( "R18_DATA".R18.Reset )
   END_RUNG wire#w3
   RUNG wire#powerrail
      I_Contact( "DI_INPUTS".R18_INPUTS_RUA.EMG_PB )
   END_RUNG wire#w4
   RUNG wire#powerrail
      Contact( "AlwaysTRUE" )
      wire#w5
      { S7_Templates := "SrcType := Int" } EQ_Contact(in1 := "Valves Data".R18_XV01.STATUS, in2 := 1)
      wire#w6
      Coil( "dummy".R18.Intl_2 )
   END_RUNG
   RUNG wire#w5
      { S7_Templates := "SrcType := Int" } EQ_Contact(in1 := "Valves Data".R18_XV03.STATUS, in2 := 1)
   END_RUNG wire#w6
   RUNG wire#w5
      { S7_Templates := "SrcType := Int" } EQ_Contact(in1 := "Valves Data".R18_XV04.STATUS, in2 := 1)
   END_RUNG wire#w6
   // the same network as SCL:
   IF "AlwaysTRUE" THEN
       #valve_R18_XV02("auto/manual" := "Valves Data"."A/M".R18,   // "valve"
                       open_auto := "R18_DATA".R18.CTS_CMD_2 OR "R18_DATA".R18.CTS_CMD_1 OR "R18_DATA".R18.CTS_CMD OR "R18_DATA".R18.CSV_CMD_3,
                       open_man := "Valves Data".R18_XV02.MCMD AND NOT "dummy".R18.Intl_2,
                       fbk_open := "A/GLR_018_XV502_OFB",
                       fbk_close := "A/GLR_018_XV502_CFB",
                       reset := "Valves Data".R18_XV02.RESET OR "R18_DATA".R18.Reset,
                       intl := NOT "DI_INPUTS".R18_INPUTS_RUA.EMG_PB,
                       Mon_En := 1,
                       mon_sp := "Valves Data".R18_XV02.MON_TIME,
                       SEMI := "Valves Data".SEMI_AUTO.R18,
                       "open/close" => "A/GLR_018_XV502_CMD",
                       FAIL_TO_OPEN => "Valves Data".R18_VALVE_FAULT.XV02_FAIL_TO_OPEN,
                       FAIL_TO_CLOSE => "Valves Data".R18_VALVE_FAULT.XV02_FAIL_TO_CLOSE,
                       status => "Valves Data".R18_XV02.STATUS);
   END_IF;
   "dummy".R18.Intl_2 := "AlwaysTRUE" AND (("Valves Data".R18_XV01.STATUS = 1) OR ("Valves Data".R18_XV03.STATUS = 1) OR ("Valves Data".R18_XV04.STATUS = 1));
END_REGION

REGION Network 189: R18_XV03
